// ---- POUs/IEC61850Server/WTURBINE/LD0/WTUR1/CDCs/FB_DO_WTURBINE_LD0_WTUR1_Beh.TcPOU
{attribute 'no_assign'}
FUNCTION_BLOCK FB_DO_WTURBINE_LD0_WTUR1_Beh EXTENDS FB_AcsiCommonDataClass
VAR_INPUT
	stVal: FB_AcsiDATypeBeh := (Fc:=ACSI_FC_ST, TrgOp:=ACSI_TrgOp_dchg OR ACSI_TrgOp_dupd, bLinkResult:=THIS^.AddDataToContainer(ipData:=stVal));
	q: FB_AcsiDATypeQuality := (Fc:=ACSI_FC_ST, TrgOp:=ACSI_TrgOp_qchg, bLinkResult:=THIS^.AddDataToContainer(ipData:=q));
	t: FB_AcsiDATypeTimeStamp := (Fc:=ACSI_FC_ST, bLinkResult:=THIS^.AddDataToContainer(ipData:=t));
END_VAR
VAR
END_VAR

END_FUNCTION_BLOCK

// ---- POUs/IEC61850Server/WTURBINE/LD0/WTUR1/CDCs/FB_DO_WTURBINE_LD0_WTUR1_TotWh.TcPOU
{attribute 'no_assign'}
FUNCTION_BLOCK FB_DO_WTURBINE_LD0_WTUR1_TotWh EXTENDS FB_AcsiCommonDataClass
VAR_INPUT
	cntVal: FB_DO_WTURBINE_LD0_WTUR1_TotWh_cntVal := (sClass:='BCR', bLinkResult:=THIS^.AddDataToContainer(ipData:=cntVal));
END_VAR
VAR
END_VAR

END_FUNCTION_BLOCK

// ---- POUs/IEC61850Server/WTURBINE/LD0/WTUR1/CDCs/FB_DO_WTURBINE_LD0_WTUR1_TotWh_cntVal.TcPOU
{attribute 'no_assign'}
FUNCTION_BLOCK FB_DO_WTURBINE_LD0_WTUR1_TotWh_cntVal EXTENDS FB_AcsiCommonDataClass
VAR_INPUT
	actVal: FB_AcsiBATypeINT64 := (Fc:=ACSI_FC_ST, TrgOp:=ACSI_TrgOp_dchg, bLinkResult:=THIS^.AddDataToContainer(ipData:=actVal));
	q: FB_AcsiDATypeQuality := (Fc:=ACSI_FC_ST, TrgOp:=ACSI_TrgOp_qchg, bLinkResult:=THIS^.AddDataToContainer(ipData:=q));
	t: FB_AcsiDATypeTimeStamp := (Fc:=ACSI_FC_ST, bLinkResult:=THIS^.AddDataToContainer(ipData:=t));
	pulsQty: FB_AcsiBATypeFLOAT32 := (Fc:=ACSI_FC_CF, TrgOp:=ACSI_TrgOp_dchg, bLinkResult:=THIS^.AddDataToContainer(ipData:=pulsQty));
END_VAR
VAR
END_VAR

END_FUNCTION_BLOCK

// ---- POUs/IEC61850Server/WTURBINE/LD0/WTUR1/CDCs/FB_DO_WTURBINE_LD0_WTUR1_TurSt.TcPOU
{attribute 'no_assign'}
FUNCTION_BLOCK FB_DO_WTURBINE_LD0_WTUR1_TurSt EXTENDS FB_AcsiCommonDataClass
VAR_INPUT
	st_: FB_DO_WTURBINE_LD0_WTUR1_TurSt_st := (sObjectName:='st', sClass:='ENS', bLinkResult:=THIS^.AddDataToContainer(ipData:=st_));
END_VAR
VAR
END_VAR

END_FUNCTION_BLOCK

// ---- POUs/IEC61850Server/WTURBINE/LD0/WTUR1/CDCs/FB_DO_WTURBINE_LD0_WTUR1_TurSt_st.TcPOU
{attribute 'no_assign'}
FUNCTION_BLOCK FB_DO_WTURBINE_LD0_WTUR1_TurSt_st EXTENDS FB_AcsiCommonDataClass
VAR_INPUT
	stVal: FB_AcsiDATypeTurSt := (Fc:=ACSI_FC_ST, TrgOp:=ACSI_TrgOp_dchg OR ACSI_TrgOp_dupd, bLinkResult:=THIS^.AddDataToContainer(ipData:=stVal));
	q: FB_AcsiDATypeQuality := (Fc:=ACSI_FC_ST, TrgOp:=ACSI_TrgOp_qchg, bLinkResult:=THIS^.AddDataToContainer(ipData:=q));
	t: FB_AcsiDATypeTimeStamp := (Fc:=ACSI_FC_ST, bLinkResult:=THIS^.AddDataToContainer(ipData:=t));
END_VAR
VAR
END_VAR

END_FUNCTION_BLOCK

// ---- POUs/IEC61850Server/WTURBINE/LD0/WTUR1/CDCs/FB_DO_WTURBINE_LD0_WTUR1_W.TcPOU
{attribute 'no_assign'}
FUNCTION_BLOCK FB_DO_WTURBINE_LD0_WTUR1_W EXTENDS FB_AcsiCommonDataClass
VAR_INPUT
	mag: FB_AcsiDATypeAnalogueValue := (Fc:=ACSI_FC_MX, TrgOp:=ACSI_TrgOp_dchg OR ACSI_TrgOp_dupd, i:=(bPresence:=FALSE), bLinkResult:=THIS^.AddDataToContainer(ipData:=mag));
	q: FB_AcsiDATypeQuality := (Fc:=ACSI_FC_MX, TrgOp:=ACSI_TrgOp_qchg, bLinkResult:=THIS^.AddDataToContainer(ipData:=q));
	t: FB_AcsiDATypeTimeStamp := (Fc:=ACSI_FC_MX, bLinkResult:=THIS^.AddDataToContainer(ipData:=t));
END_VAR
VAR
END_VAR

END_FUNCTION_BLOCK

// ---- POUs/IEC61850Server/WTURBINE/LD0/WTUR1/CDCs/FB_DO_WTURBINE_LD0_WTUR1_TurOp.TcPOU
{attribute 'no_assign'}
FUNCTION_BLOCK FB_DO_WTURBINE_LD0_WTUR1_TurOp EXTENDS FB_AcsiCommonDataClass
VAR_INPUT
	cmdAcs: FB_AcsiBATypeINT8U := (Fc:=ACSI_FC_CF, bLinkResult:=THIS^.AddDataToContainer(ipData:=cmdAcs));
	st_: FB_DO_WTURBINE_LD0_WTUR1_TurOp_st := (sObjectName:='st', sClass:='ENC', bLinkResult:=THIS^.AddDataToContainer(ipData:=st_));
END_VAR
VAR
END_VAR

END_FUNCTION_BLOCK

// ---- POUs/IEC61850Server/WTURBINE/LD0/WTUR1/CDCs/FB_DO_WTURBINE_LD0_WTUR1_TurOp_st.TcPOU
{attribute 'no_assign'}
FUNCTION_BLOCK FB_DO_WTURBINE_LD0_WTUR1_TurOp_st EXTENDS FB_AcsiCommonControllableDataClass
VAR_INPUT
	stVal: FB_AcsiDATypeTurOp := (Fc:=ACSI_FC_ST, TrgOp:=ACSI_TrgOp_dchg, bLinkResult:=THIS^.AddDataToContainer(ipData:=stVal));
	q: FB_AcsiDATypeQuality := (Fc:=ACSI_FC_ST, TrgOp:=ACSI_TrgOp_qchg, bLinkResult:=THIS^.AddDataToContainer(ipData:=q));
	t: FB_AcsiDATypeTimeStamp := (Fc:=ACSI_FC_ST, bLinkResult:=THIS^.AddDataToContainer(ipData:=t));
	ctlModel: FB_AcsiDATypeCtlModels := (Fc:=ACSI_FC_CF, TrgOp:=ACSI_TrgOp_dchg, eValue:=E_AcsiCtlModels.DirectWithNormalSecurity, bLinkResult:=THIS^.AddDataToContainer(ipData:=ctlModel));
	Cancel: FB_AcsiCDC_Cancel_ENUMERATED := (Fc:=ACSI_FC_CO, bLinkResult:=THIS^.AddDataToContainer(ipData:=Cancel));
	Oper: FB_AcsiCDC_Oper_ENUMERATED := (Fc:=ACSI_FC_CO, bLinkResult:=THIS^.AddDataToContainer(ipData:=Oper));
	SBO: FB_AcsiCDC_SBO := (Fc:=ACSI_FC_CO, bLinkResult:=THIS^.AddDataToContainer(ipData:=SBO));
	
	fbControl: FB_DirectControl := (ipCtrl:=THIS^.AddServerJob(ipEvent:=fbControl, ipCompletion:=fbControl));
END_VAR
VAR
END_VAR

END_FUNCTION_BLOCK

// ---- POUs/IEC61850Server/WTURBINE/LD0/WTUR1/CDCs/FB_DO_WTURBINE_LD0_WTUR1_DmdWSpt.TcPOU
{attribute 'no_assign'}
FUNCTION_BLOCK FB_DO_WTURBINE_LD0_WTUR1_DmdWSpt EXTENDS FB_AcsiCommonDataClass
VAR_INPUT
	val: FB_DO_WTURBINE_LD0_WTUR1_DmdWSpt_val := (sClass:='APC', bLinkResult:=THIS^.AddDataToContainer(ipData:=val));
END_VAR
VAR
END_VAR

END_FUNCTION_BLOCK

// ---- POUs/IEC61850Server/WTURBINE/LD0/WTUR1/CDCs/FB_DO_WTURBINE_LD0_WTUR1_DmdWSpt_val.TcPOU
{attribute 'no_assign'}
FUNCTION_BLOCK FB_DO_WTURBINE_LD0_WTUR1_DmdWSpt_val EXTENDS FB_AcsiCommonControllableDataClass
VAR_INPUT
	origin: FB_AcsiDATypeOriginator := (Fc:=ACSI_FC_MX, bLinkResult:=THIS^.AddDataToContainer(ipData:=origin));
	mxVal: FB_AcsiDATypeAnalogueValue := (Fc:=ACSI_FC_MX, TrgOp:=ACSI_TrgOp_dchg, i:=(bPresence:=FALSE), bLinkResult:=THIS^.AddDataToContainer(ipData:=mxVal));
	q: FB_AcsiDATypeQuality := (Fc:=ACSI_FC_MX, TrgOp:=ACSI_TrgOp_qchg, bLinkResult:=THIS^.AddDataToContainer(ipData:=q));
	t: FB_AcsiDATypeTimeStamp := (Fc:=ACSI_FC_MX, bLinkResult:=THIS^.AddDataToContainer(ipData:=t));
	ctlModel: FB_AcsiDATypeCtlModels := (Fc:=ACSI_FC_CF, TrgOp:=ACSI_TrgOp_dchg, eValue:=E_AcsiCtlModels.DirectWithNormalSecurity, bLinkResult:=THIS^.AddDataToContainer(ipData:=ctlModel));
	Oper: FB_AcsiCDC_Oper_AnalogueValue := (Fc:=ACSI_FC_CO, ctlVal:=(i:=(bPresence:=FALSE)), bLinkResult:=THIS^.AddDataToContainer(ipData:=Oper));
	SBO: FB_AcsiCDC_SBO := (Fc:=ACSI_FC_CO, bLinkResult:=THIS^.AddDataToContainer(ipData:=SBO));
	Cancel: FB_AcsiCDC_Cancel_AnalogueValue := (Fc:=ACSI_FC_CO, ctlVal:=(i:=(bPresence:=FALSE)), bLinkResult:=THIS^.AddDataToContainer(ipData:=Cancel));
	
	fbControl: FB_DirectControl := (ipCtrl:=THIS^.AddServerJob(ipEvent:=fbControl, ipCompletion:=fbControl));
// 	fbControl: FB_SboControl := (ipCtrl:=THIS^.AddServerJob(ipEvent:=fbControl, ipCompletion:=fbControl));
END_VAR
VAR
END_VAR

END_FUNCTION_BLOCK

// ---- POUs/IEC61850Server/WTURBINE/LD0/WTUR1/CDCs/FB_DO_WTURBINE_LD0_WTUR1_TurCtl.TcPOU
{attribute 'no_assign'}
FUNCTION_BLOCK FB_DO_WTURBINE_LD0_WTUR1_TurCtl EXTENDS FB_AcsiCommonDataClass
VAR_INPUT
	st_: FB_DO_WTURBINE_LD0_WTUR1_TurCtl_st := (sObjectName:='st', sClass:='ENC', bLinkResult:=THIS^.AddDataToContainer(ipData:=st_));
END_VAR
VAR
END_VAR

END_FUNCTION_BLOCK

// ---- POUs/IEC61850Server/WTURBINE/LD0/WTUR1/CDCs/FB_DO_WTURBINE_LD0_WTUR1_TurCtl_st.TcPOU
{attribute 'no_assign'}
FUNCTION_BLOCK FB_DO_WTURBINE_LD0_WTUR1_TurCtl_st EXTENDS FB_AcsiCommonControllableDataClass
VAR_INPUT
	//stVal: FB_AcsiBATypeEnumerated := (Fc:=ACSI_FC_ST, TrgOp:=ACSI_TrgOp_dchg, bLinkResult:=THIS^.AddDataToContainer(ipData:=stVal));
	stVal: FB_AcsiDATypeTurOp := (Fc:=ACSI_FC_ST, TrgOp:=ACSI_TrgOp_dchg, bLinkResult:=THIS^.AddDataToContainer(ipData:=stVal));
	q: FB_AcsiDATypeQuality := (Fc:=ACSI_FC_ST, TrgOp:=ACSI_TrgOp_qchg, bLinkResult:=THIS^.AddDataToContainer(ipData:=q));
	t: FB_AcsiDATypeTimeStamp := (Fc:=ACSI_FC_ST, bLinkResult:=THIS^.AddDataToContainer(ipData:=t));
	ctlModel: FB_AcsiDATypeCtlModels := (Fc:=ACSI_FC_CF, TrgOp:=ACSI_TrgOp_dchg, eValue:=E_AcsiCtlModels.DirectWithNormalSecurity, bLinkResult:=THIS^.AddDataToContainer(ipData:=ctlModel));
	Cancel: FB_AcsiCDC_Cancel_ENUMERATED := (Fc:=ACSI_FC_CO, bLinkResult:=THIS^.AddDataToContainer(ipData:=Cancel));
	Oper: FB_AcsiCDC_Oper_ENUMERATED := (Fc:=ACSI_FC_CO, bLinkResult:=THIS^.AddDataToContainer(ipData:=Oper));
	SBO: FB_AcsiCDC_SBO := (Fc:=ACSI_FC_CO, bLinkResult:=THIS^.AddDataToContainer(ipData:=SBO));
	
	fbControl: FB_DirectControl := (ipCtrl:=THIS^.AddServerJob(ipEvent:=fbControl, ipCompletion:=fbControl));
END_VAR
VAR
END_VAR

END_FUNCTION_BLOCK

// ---- POUs/IEC61850Server/WTURBINE/LD0/WROT1/FB_LN_WTURBINE_LD0_WROT1.TcPOU
{attribute 'no_assign'}
FUNCTION_BLOCK FB_LN_WTURBINE_LD0_WROT1 EXTENDS FB_AcsiCommonLogicalNodeClass
VAR_INPUT
	Beh: FB_DO_WTURBINE_LD0_WROT1_Beh := (sClass:='ENS', bLinkResult:=THIS^.AddDataToContainer(ipData:=Beh));
	RotSpd: FB_DO_WTURBINE_LD0_WROT1_RotSpd := (sClass:='MV', bLinkResult:=THIS^.AddDataToContainer(ipData:=RotSpd));
	BlPthAngTgt: FB_DO_WTURBINE_LD0_WROT1_BlPthAngTgt := (sClass:='MV', bLinkResult:=THIS^.AddDataToContainer(ipData:=BlPthAngTgt));
	BlPthAngVal: FB_DO_WTURBINE_LD0_WROT1_BlPthAngVal := (sClass:='MV', bLinkResult:=THIS^.AddDataToContainer(ipData:=BlPthAngVal));
END_VAR
VAR
END_VAR

END_FUNCTION_BLOCK

// ---- POUs/IEC61850Server/WTURBINE/LD0/WROT1/CDCs/FB_DO_WTURBINE_LD0_WROT1_Beh.TcPOU
{attribute 'no_assign'}
FUNCTION_BLOCK FB_DO_WTURBINE_LD0_WROT1_Beh EXTENDS FB_AcsiCommonDataClass
VAR_INPUT
	stVal: FB_AcsiDATypeBeh := (Fc:=ACSI_FC_ST, TrgOp:=ACSI_TrgOp_dchg OR ACSI_TrgOp_dupd, bLinkResult:=THIS^.AddDataToContainer(ipData:=stVal));
	q: FB_AcsiDATypeQuality := (Fc:=ACSI_FC_ST, TrgOp:=ACSI_TrgOp_qchg, bLinkResult:=THIS^.AddDataToContainer(ipData:=q));
	t: FB_AcsiDATypeTimeStamp := (Fc:=ACSI_FC_ST, bLinkResult:=THIS^.AddDataToContainer(ipData:=t));
END_VAR
VAR
END_VAR

END_FUNCTION_BLOCK

// ---- POUs/IEC61850Server/WTURBINE/LD0/WROT1/CDCs/FB_DO_WTURBINE_LD0_WROT1_RotSpd.TcPOU
{attribute 'no_assign'}
FUNCTION_BLOCK FB_DO_WTURBINE_LD0_WROT1_RotSpd EXTENDS FB_AcsiCommonDataClass
VAR_INPUT
	mag: FB_AcsiDATypeAnalogueValue := (Fc:=ACSI_FC_MX, TrgOp:=ACSI_TrgOp_dchg OR ACSI_TrgOp_dupd, i:=(bPresence:=FALSE), bLinkResult:=THIS^.AddDataToContainer(ipData:=mag));
	q: FB_AcsiDATypeQuality := (Fc:=ACSI_FC_MX, TrgOp:=ACSI_TrgOp_qchg, bLinkResult:=THIS^.AddDataToContainer(ipData:=q));
	t: FB_AcsiDATypeTimeStamp := (Fc:=ACSI_FC_MX, bLinkResult:=THIS^.AddDataToContainer(ipData:=t));
END_VAR
VAR
END_VAR

END_FUNCTION_BLOCK

// ---- POUs/IEC61850Server/WTURBINE/LD0/WROT1/CDCs/FB_DO_WTURBINE_LD0_WROT1_BlPthAngTgt.TcPOU
{attribute 'no_assign'}
FUNCTION_BLOCK FB_DO_WTURBINE_LD0_WROT1_BlPthAngTgt EXTENDS FB_AcsiCommonDataClass
VAR_INPUT
	mag: FB_AcsiDATypeAnalogueValue := (Fc:=ACSI_FC_MX, TrgOp:=ACSI_TrgOp_dchg OR ACSI_TrgOp_dupd, i:=(bPresence:=FALSE), bLinkResult:=THIS^.AddDataToContainer(ipData:=mag));
	q: FB_AcsiDATypeQuality := (Fc:=ACSI_FC_MX, TrgOp:=ACSI_TrgOp_qchg, bLinkResult:=THIS^.AddDataToContainer(ipData:=q));
	t: FB_AcsiDATypeTimeStamp := (Fc:=ACSI_FC_MX, bLinkResult:=THIS^.AddDataToContainer(ipData:=t));
END_VAR
VAR
END_VAR

END_FUNCTION_BLOCK

// ---- POUs/IEC61850Server/WTURBINE/LD0/WROT1/CDCs/FB_DO_WTURBINE_LD0_WROT1_BlPthAngVal.TcPOU
{attribute 'no_assign'}
FUNCTION_BLOCK FB_DO_WTURBINE_LD0_WROT1_BlPthAngVal EXTENDS FB_AcsiCommonDataClass
VAR_INPUT
	mag: FB_AcsiDATypeAnalogueValue := (Fc:=ACSI_FC_MX, TrgOp:=ACSI_TrgOp_dchg OR ACSI_TrgOp_dupd, i:=(bPresence:=FALSE), bLinkResult:=THIS^.AddDataToContainer(ipData:=mag));
	q: FB_AcsiDATypeQuality := (Fc:=ACSI_FC_MX, TrgOp:=ACSI_TrgOp_qchg, bLinkResult:=THIS^.AddDataToContainer(ipData:=q));
	t: FB_AcsiDATypeTimeStamp := (Fc:=ACSI_FC_MX, bLinkResult:=THIS^.AddDataToContainer(ipData:=t));
END_VAR
VAR
END_VAR

END_FUNCTION_BLOCK

// ---- POUs/IEC61850Server/WTURBINE/LD0/WCNV1/FB_LN_WTURBINE_LD0_WCNV1.TcPOU
{attribute 'no_assign'}
FUNCTION_BLOCK FB_LN_WTURBINE_LD0_WCNV1 EXTENDS FB_AcsiCommonLogicalNodeClass
VAR_INPUT
	Beh: FB_DO_WTURBINE_LD0_WCNV1_Beh := (sClass:='ENS', bLinkResult:=THIS^.AddDataToContainer(ipData:=Beh));
	Torq: FB_DO_WTURBINE_LD0_WCNV1_Torq := (sClass:='MV', bLinkResult:=THIS^.AddDataToContainer(ipData:=Torq));
END_VAR
VAR
END_VAR

END_FUNCTION_BLOCK

// ---- POUs/IEC61850Server/WTURBINE/LD0/WCNV1/CDCs/FB_DO_WTURBINE_LD0_WCNV1_Beh.TcPOU
{attribute 'no_assign'}
FUNCTION_BLOCK FB_DO_WTURBINE_LD0_WCNV1_Beh EXTENDS FB_AcsiCommonDataClass
VAR_INPUT
	stVal: FB_AcsiDATypeBeh := (Fc:=ACSI_FC_ST, TrgOp:=ACSI_TrgOp_dchg OR ACSI_TrgOp_dupd, bLinkResult:=THIS^.AddDataToContainer(ipData:=stVal));
	q: FB_AcsiDATypeQuality := (Fc:=ACSI_FC_ST, TrgOp:=ACSI_TrgOp_qchg, bLinkResult:=THIS^.AddDataToContainer(ipData:=q));
	t: FB_AcsiDATypeTimeStamp := (Fc:=ACSI_FC_ST, bLinkResult:=THIS^.AddDataToContainer(ipData:=t));
END_VAR
VAR
END_VAR

END_FUNCTION_BLOCK

// ---- POUs/IEC61850Server/WTURBINE/LD0/WCNV1/CDCs/FB_DO_WTURBINE_LD0_WCNV1_Torq.TcPOU
{attribute 'no_assign'}
FUNCTION_BLOCK FB_DO_WTURBINE_LD0_WCNV1_Torq EXTENDS FB_AcsiCommonDataClass
VAR_INPUT
	mag: FB_AcsiDATypeAnalogueValue := (Fc:=ACSI_FC_MX, TrgOp:=ACSI_TrgOp_dchg OR ACSI_TrgOp_dupd, i:=(bPresence:=FALSE), bLinkResult:=THIS^.AddDataToContainer(ipData:=mag));
	q: FB_AcsiDATypeQuality := (Fc:=ACSI_FC_MX, TrgOp:=ACSI_TrgOp_qchg, bLinkResult:=THIS^.AddDataToContainer(ipData:=q));
	t: FB_AcsiDATypeTimeStamp := (Fc:=ACSI_FC_MX, bLinkResult:=THIS^.AddDataToContainer(ipData:=t));
END_VAR
VAR
END_VAR

END_FUNCTION_BLOCK

// ---- POUs/IEC61850Server/WTURBINE/LD0/WMET1/FB_LN_WTURBINE_LD0_WMET1.TcPOU
{attribute 'no_assign'}
FUNCTION_BLOCK FB_LN_WTURBINE_LD0_WMET1 EXTENDS FB_AcsiCommonLogicalNodeClass
VAR_INPUT
	Beh: FB_DO_WTURBINE_LD0_WMET1_Beh := (sClass:='ENS', bLinkResult:=THIS^.AddDataToContainer(ipData:=Beh));
	HorWdDir: FB_DO_WTURBINE_LD0_WMET1_HorWdDir := (sClass:='MV', bLinkResult:=THIS^.AddDataToContainer(ipData:=HorWdDir));
	HorWdSpd: FB_DO_WTURBINE_LD0_WMET1_HorWdSpd := (sClass:='MV', bLinkResult:=THIS^.AddDataToContainer(ipData:=HorWdSpd));
END_VAR
VAR
END_VAR

END_FUNCTION_BLOCK

// ---- POUs/IEC61850Server/WTURBINE/LD0/WMET1/CDCs/FB_DO_WTURBINE_LD0_WMET1_Beh.TcPOU
{attribute 'no_assign'}
FUNCTION_BLOCK FB_DO_WTURBINE_LD0_WMET1_Beh EXTENDS FB_AcsiCommonDataClass
VAR_INPUT
	stVal: FB_AcsiDATypeBeh := (Fc:=ACSI_FC_ST, TrgOp:=ACSI_TrgOp_dchg OR ACSI_TrgOp_dupd, bLinkResult:=THIS^.AddDataToContainer(ipData:=stVal));
	q: FB_AcsiDATypeQuality := (Fc:=ACSI_FC_ST, TrgOp:=ACSI_TrgOp_qchg, bLinkResult:=THIS^.AddDataToContainer(ipData:=q));
	t: FB_AcsiDATypeTimeStamp := (Fc:=ACSI_FC_ST, bLinkResult:=THIS^.AddDataToContainer(ipData:=t));
END_VAR
VAR
END_VAR

END_FUNCTION_BLOCK

// ---- POUs/IEC61850Server/WTURBINE/LD0/WMET1/CDCs/FB_DO_WTURBINE_LD0_WMET1_HorWdDir.TcPOU
{attribute 'no_assign'}
FUNCTION_BLOCK FB_DO_WTURBINE_LD0_WMET1_HorWdDir EXTENDS FB_AcsiCommonDataClass
VAR_INPUT
	mag: FB_AcsiDATypeAnalogueValue := (Fc:=ACSI_FC_MX, TrgOp:=ACSI_TrgOp_dchg OR ACSI_TrgOp_dupd, i:=(bPresence:=FALSE), bLinkResult:=THIS^.AddDataToContainer(ipData:=mag));
	q: FB_AcsiDATypeQuality := (Fc:=ACSI_FC_MX, TrgOp:=ACSI_TrgOp_qchg, bLinkResult:=THIS^.AddDataToContainer(ipData:=q));
	t: FB_AcsiDATypeTimeStamp := (Fc:=ACSI_FC_MX, bLinkResult:=THIS^.AddDataToContainer(ipData:=t));
END_VAR
VAR
END_VAR

END_FUNCTION_BLOCK

// ---- POUs/IEC61850Server/WTURBINE/LD0/WMET1/CDCs/FB_DO_WTURBINE_LD0_WMET1_HorWdSpd.TcPOU
{attribute 'no_assign'}
FUNCTION_BLOCK FB_DO_WTURBINE_LD0_WMET1_HorWdSpd EXTENDS FB_AcsiCommonDataClass
VAR_INPUT
	mag: FB_AcsiDATypeAnalogueValue := (Fc:=ACSI_FC_MX, TrgOp:=ACSI_TrgOp_dchg OR ACSI_TrgOp_dupd, i:=(bPresence:=FALSE), bLinkResult:=THIS^.AddDataToContainer(ipData:=mag));
	q: FB_AcsiDATypeQuality := (Fc:=ACSI_FC_MX, TrgOp:=ACSI_TrgOp_qchg, bLinkResult:=THIS^.AddDataToContainer(ipData:=q));
	t: FB_AcsiDATypeTimeStamp := (Fc:=ACSI_FC_MX, bLinkResult:=THIS^.AddDataToContainer(ipData:=t));
END_VAR
VAR
END_VAR

END_FUNCTION_BLOCK

// ---- POUs/IEC61850Server/WTURBINE/LD0/WALM1/FB_LN_WTURBINE_LD0_WALM1.TcPOU
{attribute 'no_assign'}
FUNCTION_BLOCK FB_LN_WTURBINE_LD0_WALM1 EXTENDS FB_AcsiCommonLogicalNodeClass
VAR_INPUT
	Beh: FB_DO_WTURBINE_LD0_WALM1_Beh := (sClass:='ENS', bLinkResult:=THIS^.AddDataToContainer(ipData:=Beh));
END_VAR
VAR
END_VAR

END_FUNCTION_BLOCK

// ---- POUs/IEC61850Server/WTURBINE/LD0/WALM1/CDCs/FB_DO_WTURBINE_LD0_WALM1_Beh.TcPOU
{attribute 'no_assign'}
FUNCTION_BLOCK FB_DO_WTURBINE_LD0_WALM1_Beh EXTENDS FB_AcsiCommonDataClass
VAR_INPUT
	stVal: FB_AcsiDATypeBeh := (Fc:=ACSI_FC_ST, TrgOp:=ACSI_TrgOp_dchg OR ACSI_TrgOp_dupd, bLinkResult:=THIS^.AddDataToContainer(ipData:=stVal));
	q: FB_AcsiDATypeQuality := (Fc:=ACSI_FC_ST, TrgOp:=ACSI_TrgOp_qchg, bLinkResult:=THIS^.AddDataToContainer(ipData:=q));
	t: FB_AcsiDATypeTimeStamp := (Fc:=ACSI_FC_ST, bLinkResult:=THIS^.AddDataToContainer(ipData:=t));
END_VAR
VAR
END_VAR

END_FUNCTION_BLOCK

// ---- POUs/IEC61850Server/WTURBINE/LD0/WYAW1/FB_LN_WTURBINE_LD0_WYAW1.TcPOU
{attribute 'no_assign'}
FUNCTION_BLOCK FB_LN_WTURBINE_LD0_WYAW1 EXTENDS FB_AcsiCommonLogicalNodeClass
VAR_INPUT
	Beh: FB_DO_WTURBINE_LD0_WYAW1_Beh := (sClass:='ENS', bLinkResult:=THIS^.AddDataToContainer(ipData:=Beh));
	YwAng: FB_DO_WTURBINE_LD0_WYAW1_YwAng := (sClass:='MV', bLinkResult:=THIS^.AddDataToContainer(ipData:=YwAng));
	CabWup: FB_DO_WTURBINE_LD0_WYAW1_CabWup := (sClass:='MV', bLinkResult:=THIS^.AddDataToContainer(ipData:=CabWup));
	YwAngSpt: FB_DO_WTURBINE_LD0_WYAW1_YwAngSpt := (sClass:='SPV', bLinkResult:=THIS^.AddDataToContainer(ipData:=YwAngSpt));
END_VAR
VAR
END_VAR

END_FUNCTION_BLOCK

// ---- POUs/IEC61850Server/WTURBINE/LD0/WYAW1/CDCs/FB_DO_WTURBINE_LD0_WYAW1_Beh.TcPOU
{attribute 'no_assign'}
FUNCTION_BLOCK FB_DO_WTURBINE_LD0_WYAW1_Beh EXTENDS FB_AcsiCommonDataClass
VAR_INPUT
	stVal: FB_AcsiDATypeBeh := (Fc:=ACSI_FC_ST, TrgOp:=ACSI_TrgOp_dchg OR ACSI_TrgOp_dupd, bLinkResult:=THIS^.AddDataToContainer(ipData:=stVal));
	q: FB_AcsiDATypeQuality := (Fc:=ACSI_FC_ST, TrgOp:=ACSI_TrgOp_qchg, bLinkResult:=THIS^.AddDataToContainer(ipData:=q));
	t: FB_AcsiDATypeTimeStamp := (Fc:=ACSI_FC_ST, bLinkResult:=THIS^.AddDataToContainer(ipData:=t));
END_VAR
VAR
END_VAR

END_FUNCTION_BLOCK

// ---- POUs/IEC61850Server/WTURBINE/LD0/WYAW1/CDCs/FB_DO_WTURBINE_LD0_WYAW1_YwAng.TcPOU
{attribute 'no_assign'}
FUNCTION_BLOCK FB_DO_WTURBINE_LD0_WYAW1_YwAng EXTENDS FB_AcsiCommonDataClass
VAR_INPUT
	mag: FB_AcsiDATypeAnalogueValue := (Fc:=ACSI_FC_MX, TrgOp:=ACSI_TrgOp_dchg OR ACSI_TrgOp_dupd, i:=(bPresence:=FALSE), bLinkResult:=THIS^.AddDataToContainer(ipData:=mag));
	q: FB_AcsiDATypeQuality := (Fc:=ACSI_FC_MX, TrgOp:=ACSI_TrgOp_qchg, bLinkResult:=THIS^.AddDataToContainer(ipData:=q));
	t: FB_AcsiDATypeTimeStamp := (Fc:=ACSI_FC_MX, bLinkResult:=THIS^.AddDataToContainer(ipData:=t));
END_VAR
VAR
END_VAR

END_FUNCTION_BLOCK

// ---- POUs/IEC61850Server/WTURBINE/LD0/WYAW1/CDCs/FB_DO_WTURBINE_LD0_WYAW1_CabWup.TcPOU
{attribute 'no_assign'}
FUNCTION_BLOCK FB_DO_WTURBINE_LD0_WYAW1_CabWup EXTENDS FB_AcsiCommonDataClass
VAR_INPUT
	mag: FB_AcsiDATypeAnalogueValue := (Fc:=ACSI_FC_MX, TrgOp:=ACSI_TrgOp_dchg OR ACSI_TrgOp_dupd, i:=(bPresence:=FALSE), f:=(bPresence:=FALSE), bLinkResult:=THIS^.AddDataToContainer(ipData:=mag));
	q: FB_AcsiDATypeQuality := (Fc:=ACSI_FC_MX, TrgOp:=ACSI_TrgOp_qchg, bLinkResult:=THIS^.AddDataToContainer(ipData:=q));
	t: FB_AcsiDATypeTimeStamp := (Fc:=ACSI_FC_MX, bLinkResult:=THIS^.AddDataToContainer(ipData:=t));
END_VAR
VAR
END_VAR

END_FUNCTION_BLOCK

// ---- POUs/IEC61850Server/WTURBINE/LD0/WYAW1/CDCs/FB_DO_WTURBINE_LD0_WYAW1_YwAngSpt.TcPOU
{attribute 'no_assign'}
FUNCTION_BLOCK FB_DO_WTURBINE_LD0_WYAW1_YwAngSpt EXTENDS FB_AcsiCommonDataClass
VAR_INPUT
	val: FB_DO_WTURBINE_LD0_WYAW1_YwAngSpt_val := (sClass:='APC', bLinkResult:=THIS^.AddDataToContainer(ipData:=val));
END_VAR
VAR
END_VAR

END_FUNCTION_BLOCK

// ---- POUs/IEC61850Server/WTURBINE/LD0/WYAW1/CDCs/FB_DO_WTURBINE_LD0_WYAW1_YwAngSpt_val.TcPOU
{attribute 'no_assign'}
FUNCTION_BLOCK FB_DO_WTURBINE_LD0_WYAW1_YwAngSpt_val EXTENDS FB_AcsiCommonControllableDataClass
VAR_INPUT
	origin: FB_AcsiDATypeOriginator := (Fc:=ACSI_FC_MX, bLinkResult:=THIS^.AddDataToContainer(ipData:=origin));
	mxVal: FB_AcsiDATypeAnalogueValue := (Fc:=ACSI_FC_MX, TrgOp:=ACSI_TrgOp_dchg, i:=(bPresence:=FALSE), bLinkResult:=THIS^.AddDataToContainer(ipData:=mxVal));
	q: FB_AcsiDATypeQuality := (Fc:=ACSI_FC_MX, TrgOp:=ACSI_TrgOp_qchg, bLinkResult:=THIS^.AddDataToContainer(ipData:=q));
	t: FB_AcsiDATypeTimeStamp := (Fc:=ACSI_FC_MX, bLinkResult:=THIS^.AddDataToContainer(ipData:=t));
	ctlModel: FB_AcsiDATypeCtlModels := (Fc:=ACSI_FC_CF, TrgOp:=ACSI_TrgOp_dchg, eValue:=E_AcsiCtlModels.DirectWithNormalSecurity, bLinkResult:=THIS^.AddDataToContainer(ipData:=ctlModel));
	Oper: FB_AcsiCDC_Oper_AnalogueValue := (Fc:=ACSI_FC_CO, ctlVal:=(i:=(bPresence:=FALSE)), bLinkResult:=THIS^.AddDataToContainer(ipData:=Oper));
	
	fbControl: FB_DirectControl := (ipCtrl:=THIS^.AddServerJob(ipEvent:=fbControl, ipCompletion:=fbControl));
END_VAR
VAR
END_VAR

END_FUNCTION_BLOCK

// ---- POUs/IEC61850Server/WTURBINE/LD0/WPPD1/FB_LN_WTURBINE_LD0_WPPD1.TcPOU
{attribute 'no_assign'}
FUNCTION_BLOCK FB_LN_WTURBINE_LD0_WPPD1 EXTENDS FB_AcsiCommonLogicalNodeClass
VAR_INPUT
	Beh: FB_DO_WTURBINE_LD0_WPPD1_Beh := (sClass:='ENS', bLinkResult:=THIS^.AddDataToContainer(ipData:=Beh));
	DevSt: FB_DO_WTURBINE_LD0_WPPD1_DevSt := (sClass:='STV', bLinkResult:=THIS^.AddDataToContainer(ipData:=DevSt));
	DevOp: FB_DO_WTURBINE_LD0_WPPD1_DevOp := (sClass:='CMD', bLinkResult:=THIS^.AddDataToContainer(ipData:=DevOp));
	ClrOp: FB_DO_WTURBINE_LD0_WPPD1_ClrOp := (sClass:='CMD', bLinkResult:=THIS^.AddDataToContainer(ipData:=ClrOp));
	
	ds01: FB_DS_TEMPLATE_LD1_WPPD1_ds01 := (bLinkResult:=THIS^.AddDataSetToContainer(ipDataSet:=ds01));
	
	urcb01: FB_ScsmUrCBImplClass := (RptID:=(sValue:='WTURBINELD0/WPPD1.urcb01'), DatSet:=(sValue:='WTURBINELD0/WPPD1.ds01'), OptFlds:=(SequenceNumber:=FALSE, ReportTimeStamp:=FALSE, ReasonForInclusion:=FALSE, DataSetName:=FALSE, DataReference:=FALSE, BufferOverflow:=FALSE, EntryID:=FALSE, ConfRevision:=FALSE), TrgOps:=(DataChange:=FALSE, QualityChange:=FALSE, DataUpdate:=FALSE, Integrity:=FALSE, GeneralInterrogation:=TRUE), bLinkResult:=THIS^.AddUnbufferedReportControlBlockToContainer(ipUnbufferedReportControlBlock:=urcb01));
END_VAR
VAR
END_VAR

END_FUNCTION_BLOCK

// ---- POUs/IEC61850Server/WTURBINE/LD0/WPPD1/CDCs/FB_DO_WTURBINE_LD0_WPPD1_Beh.TcPOU
{attribute 'no_assign'}
FUNCTION_BLOCK FB_DO_WTURBINE_LD0_WPPD1_Beh EXTENDS FB_AcsiCommonDataClass
VAR_INPUT
	stVal: FB_AcsiDATypeBeh := (Fc:=ACSI_FC_ST, TrgOp:=ACSI_TrgOp_dchg OR ACSI_TrgOp_dupd, bLinkResult:=THIS^.AddDataToContainer(ipData:=stVal));
	q: FB_AcsiDATypeQuality := (Fc:=ACSI_FC_ST, TrgOp:=ACSI_TrgOp_qchg, bLinkResult:=THIS^.AddDataToContainer(ipData:=q));
	t: FB_AcsiDATypeTimeStamp := (Fc:=ACSI_FC_ST, bLinkResult:=THIS^.AddDataToContainer(ipData:=t));
END_VAR
VAR
END_VAR

END_FUNCTION_BLOCK

// ---- POUs/IEC61850Server/WTURBINE/LD0/WPPD1/CDCs/FB_DO_WTURBINE_LD0_WPPD1_DevSt.TcPOU
{attribute 'no_assign'}
FUNCTION_BLOCK FB_DO_WTURBINE_LD0_WPPD1_DevSt EXTENDS FB_AcsiCommonDataClass
VAR_INPUT
	st_: FB_DO_WTURBINE_LD0_WPPD1_DevSt_st := (sObjectName:='st', sClass:='ENS', bLinkResult:=THIS^.AddDataToContainer(ipData:=st_));
END_VAR
VAR
END_VAR

END_FUNCTION_BLOCK

// ---- POUs/IEC61850Server/WTURBINE/LD0/WPPD1/CDCs/FB_DO_WTURBINE_LD0_WPPD1_DevSt_st.TcPOU
{attribute 'no_assign'}
FUNCTION_BLOCK FB_DO_WTURBINE_LD0_WPPD1_DevSt_st EXTENDS FB_AcsiCommonDataClass
VAR_INPUT
	stVal: FB_AcsiDATypeDevSt := (Fc:=ACSI_FC_ST, TrgOp:=ACSI_TrgOp_dchg OR ACSI_TrgOp_dupd, bLinkResult:=THIS^.AddDataToContainer(ipData:=stVal));
	q: FB_AcsiDATypeQuality := (Fc:=ACSI_FC_ST, TrgOp:=ACSI_TrgOp_qchg, bLinkResult:=THIS^.AddDataToContainer(ipData:=q));
	t: FB_AcsiDATypeTimeStamp := (Fc:=ACSI_FC_ST, bLinkResult:=THIS^.AddDataToContainer(ipData:=t));
END_VAR
VAR
END_VAR

END_FUNCTION_BLOCK

// ---- POUs/IEC61850Server/WTURBINE/LD0/WPPD1/CDCs/FB_DO_WTURBINE_LD0_WPPD1_DevOp.TcPOU
{attribute 'no_assign'}
FUNCTION_BLOCK FB_DO_WTURBINE_LD0_WPPD1_DevOp EXTENDS FB_AcsiCommonDataClass
VAR_INPUT
	st_: FB_DO_WTURBINE_LD0_WPPD1_DevOp_st := (sObjectName:='st', sClass:='ENC', bLinkResult:=THIS^.AddDataToContainer(ipData:=st_));
END_VAR
VAR
END_VAR

END_FUNCTION_BLOCK

// ---- POUs/IEC61850Server/WTURBINE/LD0/WPPD1/CDCs/FB_DO_WTURBINE_LD0_WPPD1_DevOp_st.TcPOU
{attribute 'no_assign'}
FUNCTION_BLOCK FB_DO_WTURBINE_LD0_WPPD1_DevOp_st EXTENDS FB_AcsiCommonControllableDataClass
VAR_INPUT
	origin: FB_AcsiDATypeOriginator := (Fc:=ACSI_FC_ST, bLinkResult:=THIS^.AddDataToContainer(ipData:=origin));
	stVal: FB_AcsiDATypeDevOp := (Fc:=ACSI_FC_ST, TrgOp:=ACSI_TrgOp_dchg, bLinkResult:=THIS^.AddDataToContainer(ipData:=stVal));
	q: FB_AcsiDATypeQuality := (Fc:=ACSI_FC_ST, TrgOp:=ACSI_TrgOp_qchg, bLinkResult:=THIS^.AddDataToContainer(ipData:=q));
	t: FB_AcsiDATypeTimeStamp := (Fc:=ACSI_FC_ST, bLinkResult:=THIS^.AddDataToContainer(ipData:=t));
	ctlModel: FB_AcsiDATypeCtlModels := (Fc:=ACSI_FC_CF, TrgOp:=ACSI_TrgOp_dchg, bLinkResult:=THIS^.AddDataToContainer(ipData:=ctlModel));
	Cancel: FB_AcsiDATypeDelAct := (Fc:=ACSI_FC_CO, bLinkResult:=THIS^.AddDataToContainer(ipData:=Cancel));
	Oper: FB_AcsiCDC_Oper_ENUMERATED := (Fc:=ACSI_FC_CO, bLinkResult:=THIS^.AddDataToContainer(ipData:=Oper));
	SBO: FB_AcsiCDC_SBO := (Fc:=ACSI_FC_CO, bLinkResult:=THIS^.AddDataToContainer(ipData:=SBO));
	
	fbControl: FB_DirectControl := (ipCtrl:=THIS^.AddServerJob(ipEvent:=fbControl, ipCompletion:=fbControl));
END_VAR
VAR
END_VAR

END_FUNCTION_BLOCK

// ---- POUs/IEC61850Server/WTURBINE/LD0/WPPD1/CDCs/FB_DO_WTURBINE_LD0_WPPD1_ClrOp.TcPOU
{attribute 'no_assign'}
FUNCTION_BLOCK FB_DO_WTURBINE_LD0_WPPD1_ClrOp EXTENDS FB_AcsiCommonDataClass
VAR_INPUT
	st_: FB_DO_WTURBINE_LD0_WPPD1_ClrOp_st := (sObjectName:='st', sClass:='ENC', bLinkResult:=THIS^.AddDataToContainer(ipData:=st_));
END_VAR
VAR
END_VAR

END_FUNCTION_BLOCK

// ---- POUs/IEC61850Server/WTURBINE/LD0/WPPD1/CDCs/FB_DO_WTURBINE_LD0_WPPD1_ClrOp_st.TcPOU
{attribute 'no_assign'}
FUNCTION_BLOCK FB_DO_WTURBINE_LD0_WPPD1_ClrOp_st EXTENDS FB_AcsiCommonControllableDataClass
VAR_INPUT
	stVal: FB_AcsiBATypeENUMERATED := (Fc:=ACSI_FC_ST, TrgOp:=ACSI_TrgOp_dchg, bLinkResult:=THIS^.AddDataToContainer(ipData:=stVal));
	q: FB_AcsiDATypeQuality := (Fc:=ACSI_FC_ST, TrgOp:=ACSI_TrgOp_qchg, bLinkResult:=THIS^.AddDataToContainer(ipData:=q));
	t: FB_AcsiDATypeTimeStamp := (Fc:=ACSI_FC_ST, bLinkResult:=THIS^.AddDataToContainer(ipData:=t));
	ctlModel: FB_AcsiDATypeCtlModels := (Fc:=ACSI_FC_CF, TrgOp:=ACSI_TrgOp_dchg, bLinkResult:=THIS^.AddDataToContainer(ipData:=ctlModel));
	Cancel: FB_AcsiCDC_Cancel_ENUMERATED := (Fc:=ACSI_FC_CO, bLinkResult:=THIS^.AddDataToContainer(ipData:=Cancel));
	Oper: FB_AcsiCDC_Oper_ENUMERATED := (Fc:=ACSI_FC_CO, bLinkResult:=THIS^.AddDataToContainer(ipData:=Oper));
	SBO: FB_AcsiCDC_SBO := (Fc:=ACSI_FC_CO, bLinkResult:=THIS^.AddDataToContainer(ipData:=SBO));
	
	fbControl: FB_DirectControl := (ipCtrl:=THIS^.AddServerJob(ipEvent:=fbControl, ipCompletion:=fbControl));
END_VAR
VAR
END_VAR

END_FUNCTION_BLOCK

// ---- POUs/IEC61850Server/WTURBINE/LD0/WPPD1/DataSets/FB_DS_TEMPLATE_LD1_WPPD1_ds01.TcPOU
{attribute 'no_assign'}
{attribute 'call_after_init'}
FUNCTION_BLOCK FB_DS_TEMPLATE_LD1_WPPD1_ds01 EXTENDS FB_AcsiCommonDataSetClass
VAR
END_VAR

METHOD OnInit : BOOL
VAR
	nID : UDINT;
	i : UDINT;
END_VAR
// First find the nID this is part of
nID := c_nNumTurbines + 10;
FOR i := 1 TO c_nNumTurbines DO
    IF ADR(fbWTURBINE[i].WTURBINELD0.WPPD1.ds01) = ADR(THIS^) THEN
        nID := i;
        EXIT;
    END_IF
END_FOR

IF NOT DeleteAllMembers() THEN RETURN; END_IF
IF NOT AddMember(ipData:=fbWTURBINE[nID].WTURBINELD0.WYAW1.YwAng, eFc:=E_AcsiFc.MX) THEN RETURN; END_IF
IF NOT AddMember(ipData:=fbWTURBINE[nID].WTURBINELD0.WTUR1.W, eFc:=E_AcsiFc.MX) THEN RETURN; END_IF
IF NOT AddMember(ipData:=fbWTURBINE[nID].WTURBINELD0.WROT1.RotSpd, eFc:=E_AcsiFc.MX) THEN RETURN; END_IF
IF NOT AddMember(ipData:=fbWTURBINE[nID].WTURBINELD0.WROT1.BlPthAngTgt, eFc:=E_AcsiFc.MX) THEN RETURN; END_IF
IF NOT AddMember(ipData:=fbWTURBINE[nID].WTURBINELD0.WROT1.BlPthAngVal, eFc:=E_AcsiFc.MX) THEN RETURN; END_IF
IF NOT AddMember(ipData:=fbWTURBINE[nID].WTURBINELD0.WMET1.HorWdDir, eFc:=E_AcsiFc.MX) THEN RETURN; END_IF
IF NOT AddMember(ipData:=fbWTURBINE[nID].WTURBINELD0.WMET1.HorWdSpd, eFc:=E_AcsiFc.MX) THEN RETURN; END_IF
IF NOT AddMember(ipData:=fbWTURBINE[nID].WTURBINELD0.WCNV1.Torq, eFc:=E_AcsiFc.MX) THEN RETURN; END_IF
OnInit:= TRUE;
END_METHOD

END_FUNCTION_BLOCK

// ---- POUs/IEC61850Server/FB_WTURBINEServerSession.TcPOU
{attribute 'no_assign'}
FUNCTION_BLOCK FB_WTURBINEServerSession IMPLEMENTS I_ScsmAbortIndEventSink, I_ScsmAssociateIndEventSink, I_ScsmReleaseIndEventSink
VAR_INPUT
	fbConnection		: FB_iec61850ConnectionClass := (ipAbortInd:=THIS^, ipAssociateInd:=THIS^, ipReleaseInd:=THIS^);
	nID					: UDINT;
END_VAR
VAR
	_bAbort				: BOOL; (* Rising edge activates AbortReq() command execution *)
	_bDisconnect		: BOOL; (* Rising edge activates ReleaseReq() command execution *)
	
	state				: BYTE;
	eState				: E_AsyncEnvironmentState; (* Environment state *)
	eLinkStatus			: E_ScsmLinkStatus; (* Network adapter link status *)
	bBusy				: BOOL; (* If TRUE => command execution is busy *)
	bSuccess			: BOOL;
	ipResult			: I_AsyncServiceResultClass;
	sLastErrorResult	: T_MaxString;
	fbAbortReason		: FB_ServiceErrorClass := (stError:=SUCCESS_EVENT);
	sLastAbortReason	: T_MaxString;
END_VAR

fbConnection.Execute();
eState:= fbConnection.eState;
eLinkStatus:= fbConnection.eLinkStatus;

(* Execute control model control block implementations *)
// fbWTURBINE.WTURBINELD0.LLN0.Mod_.fbControl.Execute();
// fbWTURBINE.WTURBINELD0.WTUR1.CmdBlk.fbControl.Execute();
// fbWTURBINE.WTURBINELD0.WNAC1.CtlMd.fbControl.Execute();
// fbWTURBINE.WTURBINELD0.WYAW1.YwBrk.fbControl.Execute();

// fbWTURBINE[nID].WTURBINELD0.LLN0.Mod_.fbControl.Execute();
// fbWTURBINE[nID].WTURBINELD0.WTUR1.CmdBlk.fbControl.Execute();
// fbWTURBINE[nID].WTURBINELD0.WNAC1.CtlMd.fbControl.Execute();
// fbWTURBINE[nID].WTURBINELD0.WYAW1.YwBrk.fbControl.Execute();
// fbWTURBINE[nID].WTURBINELD0.WTUR1.DmdWSpt.fbControl.Execute();

(* Execute server control block implementations *)
fbWTURBINE[nID].WTURBINELD0.WPPD1.urcb01.Server.Execute();

fbWTURBINE[nID].WTURBINELD0.LLN0.Mod_.fbControl.Execute();
fbWTURBINE[nID].WTURBINELD0.WTUR1.TurOp.st_.fbControl.Execute();
fbWTURBINE[nID].WTURBINELD0.WTUR1.TurCtl.st_.fbControl.Execute();
fbWTURBINE[nID].WTURBINELD0.WTUR1.DmdWSpt.val.fbControl.Execute();
fbWTURBINE[nID].WTURBINELD0.WYAW1.YwAngSpt.val.fbControl.Execute();
fbWTURBINE[nID].WTURBINELD0.WPPD1.DevOp.st_.fbControl.Execute();
fbWTURBINE[nID].WTURBINELD0.WPPD1.ClrOp.st_.fbControl.Execute();

CASE state OF
	0: (* Initial state *)
		IF _bAbort THEN (* Abort connection => execute AbortReq() command *)
			_bAbort:= FALSE;
			bSuccess:= fbConnection.AbortReq(ipReason:=fbAbortReason, ipSink:=0, ipResult=>ipResult);
			state:= SEL(bSuccess, 100, 1);
		ELSIF eState = E_AsyncEnvironmentState.Established AND _bDisconnect THEN (* Close/release connection => execute ReleaseReq() command *)
			_bDisconnect:= FALSE;
			bSuccess:= fbConnection.ReleaseReq(ipSink:=0, ipResult=>ipResult);
			state:= SEL(bSuccess, 100, 1);
		ELSIF eState = E_AsyncEnvironmentState.Established THEN (* Connection established => exchange IED data *)
			state:= 10;
		END_IF
		_bDisconnect:= FALSE;
		(*==================================================================================================================================================================*)
	1: (* Wait for AbortReq() or ReleaseReq() command completion *)
		IF ipResult <> 0 THEN
			ipResult.Execute();
			IF NOT (bBusy:=ipResult.IsBusy()) THEN
				state:= SEL(ipResult.IsCompleted(), 100(* failed or aborted *), 0(* succeeded *));
			END_IF
		END_IF
		(*==================================================================================================================================================================*)
	10: (* connection established *)
		state:= 0;
		(*==================================================================================================================================================================*)
	100: (* Error state *)
		state:= 0;
		IF ipResult <> 0 THEN
			sLastErrorResult:= ipResult.Dump();
		END_IF
END_CASE

PROPERTY bAbort : BOOL
SET
_bAbort:= bAbort;
END_SET
END_PROPERTY

PROPERTY bDisconnect : BOOL
SET
_bDisconnect:= bDisconnect;
END_SET
END_PROPERTY

(* This method receives IEC61850::Abort.ind primitive. *)
METHOD OnAbortInd
VAR_INPUT
	ipAA		: I_ScsmAssociationClass; (* Application association. If = 0 => optional. *)
	bPAbort		: BOOL; (* TRUE => P-Abort.request(), issued by provider, FALSE => Abort.request(), issued by user. *)
	ipReason	: I_ServiceErrorClass; (* Abort reason. *)
	ipData		: I_BaseStreamClass; (* Optional data. If = 0 => default, no data. *)
END_VAR
VAR
END_VAR
IF ipReason <> 0 THEN
	sLastAbortReason:= ipReason.Dump();
END_IF
END_METHOD

(* This method receives IEC61850::Associate.ind primitive. *)
METHOD OnAssociateInd : BOOL
VAR_INPUT
	ipAA			: I_ScsmAssociationClass; (* Application association. If = 0 => optional. *)
END_VAR
VAR_OUTPUT
	ipResult		: I_AsyncServiceResultClass; (* Interface pointer to service state and result information *)
END_VAR
VAR
END_VAR
sLastAbortReason:= '';
sLastErrorResult:= '';
OnAssociateInd:= fbConnection.AssociateRsp(ipResult=>ipResult);
END_METHOD

(* This method receives IEC61850::Release.ind primitive. *)
METHOD OnReleaseInd : BOOL
VAR_INPUT
	ipAA	: I_ScsmAssociationClass; (* Application association. If = 0 => optional. *)
END_VAR
VAR_OUTPUT
	ipResult: I_AsyncServiceResultClass;
END_VAR
VAR
END_VAR
OnReleaseInd:= fbConnection.ReleaseRsp(ipResult=>ipResult);
END_METHOD

END_FUNCTION_BLOCK

// ---- POUs/IEC61850Server/FB_WTURBINEGse.TcPOU
{attribute 'no_assign'}
FUNCTION_BLOCK FB_WTURBINEGse IMPLEMENTS I_GseLinkStatusEventSink
VAR_INPUT
	fbAdapter		: FB_GseAdapterClass := (ipLinkStatus:=THIS^);
END_VAR
VAR
	eLinkStatus		: E_GseLinkStatus;
	
	bSuccess		: BOOL;
	ipError			: I_ServiceErrorClass;
	
	bStart			: BOOL := TRUE; (* Rising edge starts publishing of GOOSE data *)
	bStop			: BOOL; (* Rising edge stops publishing of GOOSE data *)
	bUpdate			: BOOL; (* Rising edge updates published GOOSE data *)
END_VAR

(*=========================================================================================*)
bSuccess:= fbAdapter.Execute(ipError=>ipError); (* Execute network adapter *)

(*=========================================================================================*)
// IF bStart THEN (* Start publishing of GOOSE data *)
// 	bStart:= FALSE;
// 	bSuccess:= fbWTURBINE.WTURBINELD0.LLN0.gocb01.Publisher.Start(ipAdapter:=fbAdapter, ipError=>ipError);
// ELSIF bStop THEN (* Stop publishing of GOOSE data *)
// 	bStop:= FALSE;
// 	bSuccess:= fbWTURBINE.WTURBINELD0.LLN0.gocb01.Publisher.Stop(ipError=>ipError);
// ELSIF bUpdate THEN (* Update published GOOSE data *)
// 	bUpdate:= FALSE;
// 	bSuccess:= fbWTURBINE.WTURBINELD0.LLN0.gocb01.Publisher.Update(ipError=>ipError);
// ELSE (* Execute publisher GoCB's *)
// 	bSuccess:= fbWTURBINE.WTURBINELD0.LLN0.gocb01.Publisher.Execute(ipError=>ipError);
// END_IF

(* This method is called every time the network adapter link status changes. *)
METHOD OnLinkStatusChange
VAR_INPUT
	ipAdapter	: I_GseAdapterClass;
	eStatus		: E_GseLinkStatus;
END_VAR
VAR
END_VAR
eLinkStatus:= eStatus;
END_METHOD

END_FUNCTION_BLOCK

// ---- POUs/IEC61850Server/FB_DirectControlEnhanced.TcPOU
FUNCTION_BLOCK FB_DirectControlEnhanced EXTENDS FB_DirectControl
VAR
END_VAR

METHOD Execute : BOOL
VAR
	bTestOk: BOOL; (*Used to cache the return value of the last '_OperativeTest' or '_DynamicTest' method call*)
	eError: E_AcsiServiceError; (*Used to cache the returned error of the last '_OperativeTest' or '_DynamicTest' method call*)
	tValue: T_UtcTime; (*Used to cache the current system time for 'tOpOk'*)
END_VAR
IF (_ipCtrl <> 0) AND_THEN (_ipCtrl.ipOper <> 0) THEN
	(* Initialize function block in the first cycle *)
	IF NOT bInit THEN
		_Init();
		bInit:=TRUE;
	END_IF

	CASE _eControlState OF
		E_DirectControlState.Ready:
			(* Check if ControlState changed in the last cycle *)
			IF bNewState THEN
				bNewState:=FALSE;
				_Reset();
			END_IF
			(* Check if a valid Oper_req was received *)
			IF bOperReq THEN
				bOperReq:=FALSE;
				(* Go to next ControlState *)
				_eControlState:=E_DirectControlState.PerformTest;
				bNewState:=TRUE;
			END_IF

		E_DirectControlState.PerformTest:
			(* Check if ControlState changed in the last cycle *)
			IF bNewState THEN
				bNewState:=FALSE;
				(* Set 'opRcvd' *)
				IF (_ipCtrl.ipOpRcvd <> 0) THEN
					_ipCtrl.ipOpRcvd.bValue:=TRUE;
				END_IF
			END_IF
			(* Trigger the operative test until it is finished *)
			IF _OperativeTest(bOperativeTestOk=>bTestOk, eError=>eError) THEN
				(* Reset 'opRcvd' *)
				IF (_ipCtrl.ipOpRcvd <> 0) THEN
					_ipCtrl.ipOpRcvd.bValue:=FALSE;
				END_IF
				IF bTestOk THEN
					(* Go to next ControlState *)
					_eControlState:=E_DirectControlState.WaitForExecution;
				ELSE
					fbCompletion.SetCompleted();
					fbCompletion.eServiceError:=eError;
					(* Go back to ControlState 'Ready' *)
					_eControlState:=E_DirectControlState.Ready;
				END_IF
				bNewState:=TRUE;
			END_IF

		E_DirectControlState.WaitForExecution:
			(* Check if ControlState changed in the last cycle *)
			IF bNewState THEN
				bNewState:=FALSE;
			END_IF
			(* Trigger the dynamic test until it is finished *)
			IF _DynamicTest(bDynamicTestOk=>bTestOk, eError=>eError) THEN
				fbCompletion.SetCompleted();
				IF bTestOk THEN
					(* Go to next ControlState *)
					IF (_ipBehVal <> 0) AND_THEN ((_ipBehVal.eValue = E_AcsiBeh.TestBlocked) OR_ELSE (_ipBehVal.eValue = E_AcsiBeh.OnBlocked)) THEN
						_eControlState:=E_DirectControlState.MirrorBlockedCommand;
					ELSE
						_eControlState:=E_DirectControlState.WaitForChange;
					END_IF
				ELSE
					fbCompletion.eServiceError:=eError;
					(* Go back to ControlState 'Ready' *)
					_eControlState:=E_DirectControlState.Ready;
				END_IF
				bNewState:=TRUE;
			END_IF

		E_DirectControlState.WaitForChange:
			(* Check if ControlState changed in the last cycle *)
			IF bNewState THEN
				bNewState:=FALSE;
				(* Set 'opOk' *)
				IF (_ipCtrl.ipOpOk <> 0) THEN
					_ipCtrl.ipOpOk.bValue:=TRUE;
				END_IF
				(* Set 'tOpOk' *)
				IF (_ipCtrl.ipTOpOk <> 0) AND_THEN (_ipCurrentAA <> 0) AND_THEN (_ipCurrentAA.GetSystemTime(tT=>tValue)) THEN
					_ipCtrl.ipTOpOk.tValue:=tValue;
				END_IF
			END_IF
			(* Update value *)
			_SetValue(uCtlVal:=_ipCtrl.ipOper.uCtlVal, ipCtlVal_AV:=_ipCtrl.ipOper.ipCtlVal_AnalogueValue);
			(* Update Timestamp 't' *)
			_UpdateTimestampValue(ipAA:=_ipCurrentAA);

			(* Reset 'opOk' *)
			IF (_ipCtrl.ipOpOk <> 0) THEN
				_ipCtrl.ipOpOk.bValue:=FALSE;
			END_IF
			(* Send CmdTerm_req+ *)
			_SendCommandTerminationReqPos(ipAA:=_ipCurrentAA, ipCtrlData:=_ipCtrl.ipOper);
			(* Go back to ControlState 'Ready' *)
			_eControlState:=E_DirectControlState.Ready;
			bNewState:=TRUE;

		E_DirectControlState.MirrorBlockedCommand:
			(* Check if ControlState changed in the last cycle *)
			IF bNewState THEN
				bNewState:=FALSE;
				(* Set 'opOk' *)
				IF (_ipCtrl.ipOpOk <> 0) THEN
					_ipCtrl.ipOpOk.bValue:=TRUE;
				END_IF
				(* Set 'tOpOk' *)
				IF (_ipCtrl.ipTOpOk <> 0) AND_THEN (_ipCurrentAA <> 0) AND_THEN (_ipCurrentAA.GetSystemTime(tT=>tValue)) THEN
					_ipCtrl.ipTOpOk.tValue:=tValue;
				END_IF
			END_IF
			(* Reset 'opOk' *)
			IF (_ipCtrl.ipOpOk <> 0) THEN
				_ipCtrl.ipOpOk.bValue:=FALSE;
			END_IF
			(* Send CmdTerm_req- *)
			_SendCommandTerminationReqNeg(ipAA:=_ipCurrentAA, ipCtrlData:=_ipCtrl.ipOper, eError:=E_AcsiApplError.NoError, ipOrigin:=_ipCtrl.ipOper.ipOrigin, ipCtlNum:=_ipCtrl.ipOper.ipCtlNum, eAddCause:=E_AcsiApplAddCause.BlockedByMode);
			(* Go back to ControlState 'Ready' *)
			_eControlState:=E_DirectControlState.Ready;
			bNewState:=TRUE;
	END_CASE
END_IF

(* Monitor transmission of LastApplError *)
CASE _nLastApplErrorReqState OF
	0:	;
	1:
		IF (_ipLastApplErrorReq <> 0) THEN
			Execute:=_ipLastApplErrorReq.Execute();
			IF NOT _ipLastApplErrorReq.IsBusy() THEN
				IF _ipLastApplErrorReq.IsCompleted() THEN
					SUPER^.SetCompleted();
				ELSE
					SUPER^.CopyFrom(ipSource:=_ipLastApplErrorReq);
				END_IF
				_nLastApplErrorReqState:=0;
			END_IF
		END_IF
END_CASE
(* Monitor transmission of CommandTermination *)
CASE _nCmdTermReqState OF
	0:	RETURN;
	1:
		IF (_ipCmdTermReq <> 0) THEN
			Execute:=_ipCmdTermReq.Execute();
			IF NOT _ipCmdTermReq.IsBusy() THEN
				IF _ipCmdTermReq.IsCompleted() THEN
					SUPER^.SetCompleted();
				ELSE
					SUPER^.CopyFrom(ipSource:=_ipLastApplErrorReq);
				END_IF
				_nCmdTermReqState:=0;
			END_IF
		END_IF
END_CASE
END_METHOD

END_FUNCTION_BLOCK

// ---- POUs/IEC61850Server/FB_SboControl.TcPOU
FUNCTION_BLOCK FB_SboControl EXTENDS FB_Control
VAR
	_eControlState: E_SboControlState; (*State of control state machine*)
	_fbSboTimer: TON; (*Timer to monitor 'sboTimeout'*)
END_VAR

(*This method is called when Cancel_req is received.
It shall check whether the Cancel request is valid and return FALSE as well as an error code if it is not.*)
METHOD PROTECTED _CheckCancelReq : BOOL
VAR_INPUT
	ipDai: I_AcsiDataAccessInfoClass; (*Additional data access info*)
END_VAR
VAR_OUTPUT
	eError: E_AcsiServiceError; (*Error code for negative response*)
END_VAR
VAR
	ipAA: I_ScsmAssociationClass; (*Interface pointer to application association*)
	stRemoteAddr: ST_SockAddr; (*Address of the client that sent the Cancel_req*)
END_VAR
IF (_ipCtrl <> 0) AND_THEN (_ipCtrl.ipCancel <> 0) THEN
	ScsmAssociation_From_Dai(in:=ipDai, out=>ipAA);
	(* Don't allow control if 'ctlModel' is set to 'status-only' *)
	IF (_ipCtrl.ipCtlModel <> 0) AND_THEN (_ipCtrl.ipCtlModel.eValue = E_AcsiCtlModels.StatusOnly) THEN
		_SendLastApplError(ipAA:=ipAA, ipCtrlData:=_ipCtrl.ipCancel, eError:=E_AcsiApplError.NoError, ipOrigin:=_ipCtrl.ipCancel.ipOrigin, ipCtlNum:=_ipCtrl.ipCancel.ipCtlNum, eAddCause:=E_AcsiApplAddCause.Unknown);
		RETURN;
	(* Cancel is always allowed in state 'Unselected' *)
	ELSIF (_eControlState = E_SboControlState.Unselected) THEN
		_CheckCancelReq:=TRUE;
		RETURN;
	(* Cancel is only allowed by the same client that sent the last accepted Sel_req *)
	ELSIF (RemoteAddress_From_ScsmAssociation(in:=ipAA, out=>stRemoteAddr)) AND_THEN (stRemoteAddr.sAddr <> _stCurrrentIp.sAddr) THEN
		_SendLastApplError(ipAA:=ipAA, ipCtrlData:=_ipCtrl.ipCancel, eError:=E_AcsiApplError.NoError, ipOrigin:=_ipCtrl.ipCancel.ipOrigin, ipCtlNum:=_ipCtrl.ipCancel.ipCtlNum, eAddCause:=E_AcsiApplAddCause.LockedByOtherClient);
		RETURN;
	(* Cancel is not allowed in state 'Operate' *)
	ELSIF (_eControlState = E_SboControlState.Operate) THEN
		_SendLastApplError(ipAA:=ipAA, ipCtrlData:=_ipCtrl.ipCancel, eError:=E_AcsiApplError.NoError, ipOrigin:=_ipCtrl.ipCancel.ipOrigin, ipCtlNum:=_ipCtrl.ipCancel.ipCtlNum, eAddCause:=E_AcsiApplAddCause.CommandAlreadyInExecution);
		RETURN;
	(* Cancel is valid *)
	ELSE
		_CheckCancelReq:=TRUE;
	END_IF
END_IF
END_METHOD

//Resets all local values
METHOD PROTECTED _Reset
VAR
END_VAR
SUPER^._Reset();
(* Reset timer *)
_fbSboTimer(IN:=FALSE);
END_METHOD

METHOD Execute : BOOL
VAR
	bTestOk: BOOL; (*Used to cache the return value of the last '_OperativeTest' or '_DynamicTest' method call*)
	eError: E_AcsiServiceError; (*Used to cache the returned error of the last '_OperativeTest' or '_DynamicTest' method call*)
	tValue: T_UtcTime; (*Used to cache the current system time for 'tOpOk'*)
END_VAR
IF (_ipCtrl <> 0) AND_THEN (_ipCtrl.ipOper <> 0) THEN
	(* Initialize function block in the first cycle *)
	IF NOT bInit THEN
		_Init();
		bInit:=TRUE;
	END_IF

	CASE _eControlState OF
		E_SboControlState.Unselected:
			(* Check if ControlState changed in the last cycle *)
			IF bNewState THEN
				bNewState:=FALSE;
				_Reset();
				(* Reset 'stSeld' *)
				IF (_ipCtrl.ipStSeld <> 0) THEN
					_ipCtrl.ipStSeld.bValue:=FALSE;
				END_IF
			END_IF
			(* Check if a valid Cancel_req was received *)
			IF bCancelReq THEN
				bCancelReq:=FALSE;
			END_IF
			(* Check if a valid Sel_req was received *)
			IF bSelReq THEN
				bSelReq:=FALSE;
				(* Set 'stSeld' *)
				IF (_ipCtrl.ipStSeld <> 0) THEN
					_ipCtrl.ipStSeld.bValue:=TRUE;
				END_IF
				(* Go to next ControlState *)
				_eControlState:=E_SboControlState.Ready;
				bNewState:=TRUE;
			END_IF

		E_SboControlState.Ready:
			(* Check if ControlState changed in the last cycle *)
			IF bNewState THEN
				bNewState:=FALSE;
				(* Start timer *)
				IF (_ipCtrl.ipSboTimeout <> 0) THEN
					_fbSboTimer(IN:=TRUE, PT:=DWORD_TO_TIME(_ipCtrl.ipSboTimeout.nValue));
				END_IF
			END_IF
			_fbSboTimer();
			(* Check if a valid Cancel_req was received, 'sboTimeout' was exceeded or the association was lost *)
			IF bCancelReq OR_ELSE _fbSboTimer.Q OR_ELSE ((_ipCurrentAA <> 0) AND_THEN (_ipCurrentAA.eState <> E_AsyncEnvironmentState.Established)) THEN
				bCancelReq:=FALSE;
				_fbSboTimer(IN:=FALSE);
				(* Go to next ControlState *)
				_eControlState:=E_SboControlState.EndSelection;
				bNewState:=TRUE;
			END_IF
			(* Check if a valid Oper_req was received *)
			IF bOperReq THEN
				bOperReq:=FALSE;
				(* Go to next ControlState *)
				_eControlState:=E_SboControlState.PerformTest;
				bNewState:=TRUE;
			END_IF

		E_SboControlState.PerformTest:
			(* Check if ControlState changed in the last cycle *)
			IF bNewState THEN
				bNewState:=FALSE;
				(* Set 'opRcvd' *)
				IF (_ipCtrl.ipOpRcvd <> 0) THEN
					_ipCtrl.ipOpRcvd.bValue:=TRUE;
				END_IF
			END_IF
			(* Check if a valid Cancel_req was received *)
			IF bCancelReq THEN
				bCancelReq:=FALSE;
				(* Send Oper_resp- *)
				_SendLastApplError(ipAA:=_ipCurrentAA, ipCtrlData:=_ipCtrl.ipOper, eError:=E_AcsiApplError.NoError, ipOrigin:=_ipCtrl.ipOper.ipOrigin, ipCtlNum:=_ipCtrl.ipOper.ipCtlNum, eAddCause:=E_AcsiApplAddCause.AbortionByCancel);
				fbOperCompletion.SetCompleted();
				fbOperCompletion.eServiceError:=E_AcsiServiceError.AccessViolation;
				(* Go to ControlState 'EndSelection' *)
				_eControlState:=E_SboControlState.EndSelection;
				bNewState:=TRUE;
			END_IF
			(* Trigger the operative test until it is finished *)
			IF _OperativeTest(bOperativeTestOk=>bTestOk, eError=>eError) THEN
				(* Reset 'opRcvd' *)
				IF (_ipCtrl.ipOpRcvd <> 0) THEN
					_ipCtrl.ipOpRcvd.bValue:=FALSE;
				END_IF
				IF bTestOk THEN
					(* Go to next ControlState *)
					_eControlState:=E_SboControlState.WaitForExecution;
				ELSE
					fbOperCompletion.SetCompleted();
					fbOperCompletion.eServiceError:=eError;
					(* Go to ControlState 'EndSelection' *)
					_eControlState:=E_SboControlState.EndSelection;
				END_IF
				bNewState:=TRUE;
			END_IF

		E_SboControlState.WaitForExecution:
			(* Check if ControlState changed in the last cycle *)
			IF bNewState THEN
				bNewState:=FALSE;
			END_IF
			(* Check if a Cancel_req was received *)
			IF bCancelReq THEN
				bCancelReq:=FALSE;
				(* Send Oper_resp- *)
				_SendLastApplError(ipAA:=_ipCurrentAA, ipCtrlData:=_ipCtrl.ipOper, eError:=E_AcsiApplError.NoError, ipOrigin:=_ipCtrl.ipOper.ipOrigin, ipCtlNum:=_ipCtrl.ipOper.ipCtlNum, eAddCause:=E_AcsiApplAddCause.AbortionByCancel);
				fbOperCompletion.SetCompleted();
				fbOperCompletion.eServiceError:=E_AcsiServiceError.AccessViolation;
				(* Go to ControlState 'EndSelection' *)
				_eControlState:=E_SboControlState.EndSelection;
				bNewState:=TRUE;
			END_IF
			(* Trigger the dynamic test until it is finished *)
			IF _DynamicTest(bDynamicTestOk=>bTestOk, eError=>eError) THEN
				fbOperCompletion.SetCompleted();
				IF bTestOk THEN
					(* Go to next ControlState *)
					IF (_ipBehVal <> 0) AND_THEN ((_ipBehVal.eValue = E_AcsiBeh.TestBlocked) OR_ELSE (_ipBehVal.eValue = E_AcsiBeh.OnBlocked)) THEN
						_eControlState:=E_SboControlState.MirrorBlockedCommand;
					ELSE
						_eControlState:=E_SboControlState.Operate;
					END_IF
				ELSE
					fbOperCompletion.eServiceError:=eError;
					(* Go to ControlState 'EndSelection' *)
					_eControlState:=E_SboControlState.EndSelection;
				END_IF
				bNewState:=TRUE;
			END_IF

		E_SboControlState.Operate:
			(* Check if ControlState changed in the last cycle *)
			IF bNewState THEN
				bNewState:=FALSE;
				(* Set 'opOk' *)
				IF (_ipCtrl.ipOpOk <> 0) THEN
					_ipCtrl.ipOpOk.bValue:=TRUE;
				END_IF
				(* Set 'tOpOk' *)
				IF (_ipCtrl.ipTOpOk <> 0) AND_THEN (_ipCurrentAA <> 0) AND_THEN (_ipCurrentAA.GetSystemTime(tT=>tValue)) THEN
					_ipCtrl.ipTOpOk.tValue:=tValue;
				END_IF
			END_IF
			(* Update value *)
			_SetValue(uCtlVal:=_ipCtrl.ipOper.uCtlVal, ipCtlVal_AV:=_ipCtrl.ipOper.ipCtlVal_AnalogueValue);
			(* Update Timestamp 't' *)
			_UpdateTimestampValue(ipAA:=_ipCurrentAA);

			(* Reset 'opOk' *)
			IF (_ipCtrl.ipOpOk <> 0) THEN
				_ipCtrl.ipOpOk.bValue:=FALSE;
			END_IF
			(* Go to next ControlState *)
			IF (_ipCtrl.ipSboClass <> 0) AND_THEN (_ipCtrl.ipSboClass.eValue = E_AcsiSboClasses.OperateMany) THEN
				_eControlState:=E_SboControlState.Ready;
			ELSE
				_eControlState:=E_SboControlState.EndSelection;
			END_IF
			bNewState:=TRUE;

		E_SboControlState.MirrorBlockedCommand:
			(* Check if ControlState changed in the last cycle *)
			IF bNewState THEN
				bNewState:=FALSE;
				(* Set 'opOk' *)
				IF (_ipCtrl.ipOpOk <> 0) THEN
					_ipCtrl.ipOpOk.bValue:=TRUE;
				END_IF
				(* Set 'tOpOk' *)
				IF (_ipCtrl.ipTOpOk <> 0) AND_THEN (_ipCurrentAA <> 0) AND_THEN (_ipCurrentAA.GetSystemTime(tT=>tValue)) THEN
					_ipCtrl.ipTOpOk.tValue:=tValue;
				END_IF
			END_IF
			(* Reset 'opOk' *)
			IF (_ipCtrl.ipOpOk <> 0) THEN
				_ipCtrl.ipOpOk.bValue:=FALSE;
			END_IF
			(* Go to next ControlState *)
			IF (_ipCtrl.ipSboClass <> 0) AND_THEN (_ipCtrl.ipSboClass.eValue = E_AcsiSboClasses.OperateMany) THEN
				_eControlState:=E_SboControlState.Ready;
			ELSE
				_eControlState:=E_SboControlState.EndSelection;
			END_IF
			bNewState:=TRUE;

		E_SboControlState.EndSelection:
			(* Check if ControlState changed in the last cycle *)
			IF bNewState THEN
				bNewState:=FALSE;
				(* Reset 'stSeld' *)
				IF (_ipCtrl.ipStSeld <> 0) THEN
					_ipCtrl.ipStSeld.bValue:=FALSE;
				END_IF
			END_IF
			(* Go to next ControlState *)
			_eControlState:=E_SboControlState.Unselected;
			bNewState:=TRUE;
	END_CASE
END_IF

(* Monitor transmission of LastApplError *)
CASE _nLastApplErrorReqState OF
	0:	RETURN;
	1:
		IF (_ipLastApplErrorReq <> 0) THEN
			Execute:=_ipLastApplErrorReq.Execute();
			IF NOT _ipLastApplErrorReq.IsBusy() THEN
				IF _ipLastApplErrorReq.IsCompleted() THEN
					SUPER^.SetCompleted();
				ELSE
					SUPER^.CopyFrom(ipSource:=_ipLastApplErrorReq);
				END_IF
				_nLastApplErrorReqState:=0;
			END_IF
		END_IF
END_CASE
END_METHOD

METHOD OnCompletionWaitEvent : BOOL
VAR_INPUT
	ipDai: I_AcsiDataAccessInfoClass;
	ipData: I_AcsiCommonDataClass;
	eFc: E_AcsiFc;
END_VAR
VAR_OUTPUT
	ipResult: I_AcsiServiceResultClass := fbCompletion;
END_VAR
VAR
	eServiceError: E_AcsiServiceError;
	ipAA: I_ScsmAssociationClass; (*Interface pointer to application association*)
END_VAR
fbCompletion.SetCompleted();
IF (ipDai = 0) OR_ELSE (ipData = 0) THEN
	fbCompletion.eServiceError:=E_AcsiServiceError.AccessViolation;
	RETURN;
END_IF

(* Check if an Operate request is received *)
IF (ipDai.eService = E_AcsiServiceType.SetDataValues) THEN
	IF	(ipData.sObjectName = 'Oper') THEN
		ScsmAssociation_From_Dai(in:=ipDai, out=>_ipCurrentAA);
		fbOperCompletion.SetBusy();
		ipResult:=fbOperCompletion;
		bOperReq:=TRUE;
		OnCompletionWaitEvent:=TRUE;
	ELSIF (ipData.sObjectName = 'Cancel') THEN
		fbCancelCompletion.SetCompleted();
		ipResult:=fbCancelCompletion;
		IF _CheckCancelReq(ipDai:=ipDai, eError=>eServiceError) THEN
			bCancelReq:=TRUE;
		ELSE
			fbCancelCompletion.eServiceError:=eServiceError;
		END_IF
	END_IF
END_IF
END_METHOD

(*Implementation of user application data update event method.*)
METHOD OnGetVEvent
VAR_INPUT
	ipDai: I_AcsiDataAccessInfoClass; (*Additional data access info*)
	ipData: I_AcsiCommonDataClass; (*Interface pointer to data object*)
	eFc: E_AcsiFc; (*Functional constraint*)
END_VAR
VAR
END_VAR
IF (eFc = E_AcsiFc.CO) AND_THEN (_ipCtrl <> 0) AND_THEN (ipDai <> 0) AND_THEN (ipDai.Read) AND_THEN (ipDai.ipAccessData <> 0) THEN
	IF (ipDai.ipAccessData.sObjectName = 'SBO') AND_THEN (_ipCtrl.ipSBO <> 0) THEN
		(* Reset value of 'SBO' *)
		_ipCtrl.ipSBO.sValue:='';
	END_IF
END_IF
END_METHOD

(*Implementation of user application data update event method.*)
METHOD OnGetVPreEvent : E_AcsiServiceError
VAR_INPUT
	ipDai: I_AcsiDataAccessInfoClass; (*Additional data access info*)
	ipData: I_AcsiCommonDataClass; (*Interface pointer to data object*)
	eFc: E_AcsiFc; (*Functional constraint*)
END_VAR
VAR
END_VAR
IF (eFc = E_AcsiFc.CO) AND_THEN (_ipCtrl <> 0) AND_THEN (ipDai <> 0) AND_THEN (ipDai.Read) AND_THEN (ipDai.ipAccessData <> 0) THEN
	IF (ipDai.ipAccessData.sObjectName = 'SBO') AND_THEN (_ipCtrl.ipSBO <> 0) THEN
		(* Only allow 'Select' requests in state 'Unselected' *)
		IF (_eControlState = E_SboControlState.Unselected) THEN
			_ipCtrl.ipSBO.sValue:=_ipCtrl.ipSBO.GetSboReference();
			bSelReq:=TRUE;
		ELSE
			_ipCtrl.ipSBO.sValue:='';
		END_IF
	END_IF
END_IF
END_METHOD

(*Implementation of user application data update event method.*)
METHOD OnSetVPreEvent : E_AcsiServiceError
VAR_INPUT
	ipDai: I_AcsiDataAccessInfoClass; (*Additional data access info*)
	ipMemory: I_AnyMemoryBuffer; (*Interface pointer to buffer containig new value data*)
	ipData: I_AcsiCommonDataClass; (*Interface pointer to data object*)
	eFc: E_AcsiFc; (*Functional constraint*)
END_VAR
VAR_OUTPUT
	ipLastApplError: I_AcsiDATypeLastApplError; (*IF <> 0 => send LastApplError request*)
END_VAR
VAR
	ipAA: I_ScsmAssociationClass; (*Interface pointer to application association*)
	bItself: BOOL; (*If TRUE => Checking object is sub-data object itself*)
END_VAR
IF (eFc = E_AcsiFc.CO) AND_THEN (_ipCtrl <> 0) AND_THEN (ipDai <> 0) AND_THEN (ipDai.Write) AND_THEN (ipDai.ipAccessData <> 0) AND_THEN (ipData <> 0) AND_THEN ScsmAssociation_From_Dai(in:=ipDai, out=>ipAA) THEN
	IF (_ipCtrl.ipOper <> 0) AND_THEN (_ipCtrl.ipOper.ipOrigin <> 0) AND_THEN (_ipCtrl.ipOper.ipCtlNum <> 0) THEN
		(* Check for invalid write attemps to prevent 'Oper' from being overwritten while a control request is being executed *)
		IF (ipDai.ipAccessData.sObjectName = 'Oper') THEN
			(* Only allow 'Oper' requests in state 'Ready' *)
			IF (_eControlState <> E_SboControlState.Ready) THEN
				ipLastApplError:=ipAA.SetAdditionalCauseDiag(ipCtrlData:=_ipCtrl.ipOper, eError:=E_AcsiApplError.NoError, stOrigin:=_ipCtrl.ipOper.ipOrigin.stOrigin, nCtlNum:=_ipCtrl.ipOper.ipCtlNum.nValue, eAddCause:=E_AcsiApplAddCause.CommandAlreadyInExecution);
				OnSetVPreEvent:=E_AcsiServiceError.AccessViolation;
				RETURN;
			END_IF
		ELSIF (_ipCtrl.ipOper.HasDataSubObject(ipData:=ipDai.ipAccessData, bItself=>bItself) AND_THEN (NOT bItself)) THEN
			(* Don't allow write access to subdata of 'Oper'*)
			ipLastApplError:=ipAA.SetAdditionalCauseDiag(ipCtrlData:=_ipCtrl.ipOper, eError:=E_AcsiApplError.NoError, stOrigin:=_ipCtrl.ipOper.ipOrigin.stOrigin, nCtlNum:=_ipCtrl.ipOper.ipCtlNum.nValue, eAddCause:=E_AcsiApplAddCause.NotSupported);
			OnSetVPreEvent:=E_AcsiServiceError.AccessViolation;
			RETURN;
		END_IF
	END_IF
	IF (_ipCtrl.ipCancel <> 0) AND_THEN (_ipCtrl.ipCancel.ipOrigin <> 0) AND_THEN (_ipCtrl.ipCancel.ipCtlNum <> 0) THEN
		IF (ipDai.ipAccessData.sObjectName <> 'Cancel') AND_THEN (_ipCtrl.ipCancel.HasDataSubObject(ipData:=ipDai.ipAccessData)) THEN
			(* Don't allow write access to subdata of 'Cancel'*)
			ipLastApplError:=ipAA.SetAdditionalCauseDiag(ipCtrlData:=_ipCtrl.ipCancel, eError:=E_AcsiApplError.NoError, stOrigin:=_ipCtrl.ipCancel.ipOrigin.stOrigin, nCtlNum:=_ipCtrl.ipCancel.ipCtlNum.nValue, eAddCause:=E_AcsiApplAddCause.NotSupported);
			OnSetVPreEvent:=E_AcsiServiceError.AccessViolation;
			RETURN;
		END_IF
	END_IF
	IF (ipData.sObjectName = 'SBO') THEN
		(* Don't allow write access to 'SBO'*)
		OnSetVPreEvent:=E_AcsiServiceError.AccessViolation;
		RETURN;
	END_IF
END_IF
END_METHOD

END_FUNCTION_BLOCK

// ---- POUs/IEC61850Server/FB_SboControlEnhanced.TcPOU
FUNCTION_BLOCK FB_SboControlEnhanced EXTENDS FB_SboControl
VAR
END_VAR

METHOD Execute : BOOL
VAR
	bTestOk: BOOL; (*Used to cache the return value of the last '_OperativeTest' or '_DynamicTest' method call*)
	eError: E_AcsiServiceError; (*Used to cache the returned error of the last '_OperativeTest' or '_DynamicTest' method call*)
	tValue: T_UtcTime; (*Used to cache the current system time for 'tOpOk'*)
END_VAR
IF (_ipCtrl <> 0) AND_THEN (_ipCtrl.ipOper <> 0) THEN
	(* Initialize function block in the first cycle *)
	IF NOT bInit THEN
		_Init();
		bInit:=TRUE;
	END_IF

	CASE _eControlState OF
		E_SboControlState.Unselected:
			(* Check if ControlState changed in the last cycle *)
			IF bNewState THEN
				bNewState:=FALSE;
				_Reset();
			END_IF
			(* Check if a valid Cancel_req was received *)
			IF bCancelReq THEN
				bCancelReq:=FALSE;
			END_IF
			(* Check if a valid SelVal_req was received *)
			IF bSelValReq THEN
				bSelValReq:=FALSE;
				(* Go to next ControlState *)
				_eControlState:=E_SboControlState.Select_PerformTest;
				bNewState:=TRUE;
			END_IF

		E_SboControlState.Select_PerformTest:
			(* Check if ControlState changed in the last cycle *)
			IF bNewState THEN
				bNewState:=FALSE;
			END_IF
			(* Trigger the test until it is finished *)
			IF _Test(bTestOk=>bTestOk, eError=>eError) THEN
				IF bTestOk THEN
					(* Go to next ControlState *)
					_eControlState:=E_SboControlState.WaitForSelection;
				ELSE
					fbSelValCompletion.SetCompleted();
					fbSelValCompletion.eServiceError:=eError;
					(* Go back to ControlState 'Unselected' *)
					_eControlState:=E_SboControlState.Unselected;
				END_IF
				bNewState:=TRUE;
			END_IF

		E_SboControlState.WaitForSelection:
			(* Check if ControlState changed in the last cycle *)
			IF bNewState THEN
				bNewState:=FALSE;
			END_IF
			(* Set 'stSeld' *)
			IF (_ipCtrl.ipStSeld <> 0) THEN
				_ipCtrl.ipStSeld.bValue:=TRUE;
			END_IF
			fbSelValCompletion.SetCompleted();
			(* Go to next ControlState *)
			_eControlState:=E_SboControlState.Ready;
			bNewState:=TRUE;

		E_SboControlState.Ready:
			(* Check if ControlState changed in the last cycle *)
			IF bNewState THEN
				bNewState:=FALSE;
				(* Start timer *)
				IF (_ipCtrl.ipSboTimeout <> 0) THEN
					_fbSboTimer(IN:=TRUE, PT:=DWORD_TO_TIME(_ipCtrl.ipSboTimeout.nValue));
				END_IF
			END_IF
			_fbSboTimer();
			(* Check if a valid Cancel_req was received, 'sboTimeout' was exceeded or the association was lost *)
			IF bCancelReq OR_ELSE _fbSboTimer.Q OR_ELSE ((_ipCurrentAA <> 0) AND_THEN (_ipCurrentAA.eState <> E_AsyncEnvironmentState.Established)) THEN
				bCancelReq:=FALSE;
				_fbSboTimer(IN:=FALSE);
				(* Go to next ControlState *)
				_eControlState:=E_SboControlState.EndSelection;
				bNewState:=TRUE;
			END_IF
			(* Check if a valid Oper_req was received *)
			IF bOperReq THEN
				bOperReq:=FALSE;
				(* Go to next ControlState *)
				_eControlState:=E_SboControlState.PerformTest;
				bNewState:=TRUE;
			END_IF

		E_SboControlState.PerformTest:
			(* Check if ControlState changed in the last cycle *)
			IF bNewState THEN
				bNewState:=FALSE;
				(* Set 'opRcvd' *)
				IF (_ipCtrl.ipOpRcvd <> 0) THEN
					_ipCtrl.ipOpRcvd.bValue:=TRUE;
				END_IF
			END_IF
			(* Check if a valid Cancel_req was received *)
			IF bCancelReq THEN
				bCancelReq:=FALSE;
				(* Send Oper_resp- *)
				_SendLastApplError(ipAA:=_ipCurrentAA, ipCtrlData:=_ipCtrl.ipOper, eError:=E_AcsiApplError.NoError, ipOrigin:=_ipCtrl.ipOper.ipOrigin, ipCtlNum:=_ipCtrl.ipOper.ipCtlNum, eAddCause:=E_AcsiApplAddCause.AbortionByCancel);
				fbOperCompletion.SetCompleted();
				fbOperCompletion.eServiceError:=E_AcsiServiceError.AccessViolation;
				(* Go to ControlState 'EndSelection' *)
				_eControlState:=E_SboControlState.EndSelection;
				bNewState:=TRUE;
			END_IF
			(* Trigger the operative test until it is finished *)
			IF _OperativeTest(bOperativeTestOk=>bTestOk, eError=>eError) THEN
				(* Reset 'opRcvd' *)
				IF (_ipCtrl.ipOpRcvd <> 0) THEN
					_ipCtrl.ipOpRcvd.bValue:=FALSE;
				END_IF
				IF bTestOk THEN
					(* Go to next ControlState *)
					_eControlState:=E_SboControlState.WaitForExecution;
				ELSE
					fbOperCompletion.SetCompleted();
					fbOperCompletion.eServiceError:=eError;
					(* Go to ControlState 'EndSelection' *)
					_eControlState:=E_SboControlState.EndSelection;
				END_IF
				bNewState:=TRUE;
			END_IF

		E_SboControlState.WaitForExecution:
			(* Check if ControlState changed in the last cycle *)
			IF bNewState THEN
				bNewState:=FALSE;
			END_IF
			(* Check if a Cancel_req was received *)
			IF bCancelReq THEN
				bCancelReq:=FALSE;
				(* Send Oper_resp- *)
				_SendLastApplError(ipAA:=_ipCurrentAA, ipCtrlData:=_ipCtrl.ipOper, eError:=E_AcsiApplError.NoError, ipOrigin:=_ipCtrl.ipOper.ipOrigin, ipCtlNum:=_ipCtrl.ipOper.ipCtlNum, eAddCause:=E_AcsiApplAddCause.AbortionByCancel);
				fbOperCompletion.SetCompleted();
				fbOperCompletion.eServiceError:=E_AcsiServiceError.AccessViolation;
				(* Go to ControlState 'EndSelection' *)
				_eControlState:=E_SboControlState.EndSelection;
				bNewState:=TRUE;
			END_IF
			(* Trigger the dynamic test until it is finished *)
			IF _DynamicTest(bDynamicTestOk=>bTestOk, eError=>eError) THEN
				fbOperCompletion.SetCompleted();
				IF bTestOk THEN
					(* Go to next ControlState *)
					IF (_ipBehVal <> 0) AND_THEN ((_ipBehVal.eValue = E_AcsiBeh.TestBlocked) OR_ELSE (_ipBehVal.eValue = E_AcsiBeh.OnBlocked)) THEN
						_eControlState:=E_SboControlState.MirrorBlockedCommand;
					ELSE
						_eControlState:=E_SboControlState.WaitForChange;
					END_IF
				ELSE
					fbOperCompletion.eServiceError:=eError;
					(* Go to ControlState 'EndSelection' *)
					_eControlState:=E_SboControlState.EndSelection;
				END_IF
				bNewState:=TRUE;
			END_IF

		E_SboControlState.WaitForChange:
			(* Check if ControlState changed in the last cycle *)
			IF bNewState THEN
				bNewState:=FALSE;
				(* Set 'opOk' *)
				IF (_ipCtrl.ipOpOk <> 0) THEN
					_ipCtrl.ipOpOk.bValue:=TRUE;
				END_IF
				(* Set 'tOpOk' *)
				IF (_ipCtrl.ipTOpOk <> 0) AND_THEN (_ipCurrentAA <> 0) AND_THEN (_ipCurrentAA.GetSystemTime(tT=>tValue)) THEN
					_ipCtrl.ipTOpOk.tValue:=tValue;
				END_IF
			END_IF
			(* Update value *)
			_SetValue(uCtlVal:=_ipCtrl.ipOper.uCtlVal, ipCtlVal_AV:=_ipCtrl.ipOper.ipCtlVal_AnalogueValue);
			(* Update Timestamp 't' *)
			_UpdateTimestampValue(ipAA:=_ipCurrentAA);

			(* Reset 'opOk' *)
			IF (_ipCtrl.ipOpOk <> 0) THEN
				_ipCtrl.ipOpOk.bValue:=FALSE;
			END_IF
			(* Send CmdTerm_req+ *)
			_SendCommandTerminationReqPos(ipAA:=_ipCurrentAA, ipCtrlData:=_ipCtrl.ipOper);
			(* Go to next ControlState *)
			IF (_ipCtrl.ipSboClass <> 0) AND_THEN (_ipCtrl.ipSboClass.eValue = E_AcsiSboClasses.OperateMany) THEN
				_eControlState:=E_SboControlState.Ready;
			ELSE
				_eControlState:=E_SboControlState.EndSelection;
			END_IF
			bNewState:=TRUE;

		E_SboControlState.MirrorBlockedCommand:
			(* Check if ControlState changed in the last cycle *)
			IF bNewState THEN
				bNewState:=FALSE;
				(* Set 'opOk' *)
				IF (_ipCtrl.ipOpOk <> 0) THEN
					_ipCtrl.ipOpOk.bValue:=TRUE;
				END_IF
				(* Set 'tOpOk' *)
				IF (_ipCtrl.ipTOpOk <> 0) AND_THEN (_ipCurrentAA <> 0) AND_THEN (_ipCurrentAA.GetSystemTime(tT=>tValue)) THEN
					_ipCtrl.ipTOpOk.tValue:=tValue;
				END_IF
			END_IF
			(* Reset 'opOk' *)
			IF (_ipCtrl.ipOpOk <> 0) THEN
				_ipCtrl.ipOpOk.bValue:=FALSE;
			END_IF
			(* Send CmdTerm_req- *)
			_SendCommandTerminationReqNeg(ipAA:=_ipCurrentAA, ipCtrlData:=_ipCtrl.ipOper, eError:=E_AcsiApplError.NoError, ipOrigin:=_ipCtrl.ipOper.ipOrigin, ipCtlNum:=_ipCtrl.ipOper.ipCtlNum, eAddCause:=E_AcsiApplAddCause.BlockedByMode);
			(* Go to next ControlState *)
			IF (_ipCtrl.ipSboClass <> 0) AND_THEN (_ipCtrl.ipSboClass.eValue = E_AcsiSboClasses.OperateMany) THEN
				_eControlState:=E_SboControlState.Ready;
			ELSE
				_eControlState:=E_SboControlState.EndSelection;
			END_IF
			bNewState:=TRUE;

		E_SboControlState.EndSelection:
			(* Check if ControlState changed in the last cycle *)
			IF bNewState THEN
				bNewState:=FALSE;
				(* Reset 'stSeld' *)
				IF (_ipCtrl.ipStSeld <> 0) THEN
					_ipCtrl.ipStSeld.bValue:=FALSE;
				END_IF
			END_IF
			(* Go to next ControlState *)
			_eControlState:=E_SboControlState.Unselected;
			bNewState:=TRUE;
	END_CASE
END_IF

(* Monitor transmission of LastApplError *)
CASE _nLastApplErrorReqState OF
	0:	;
	1:
		IF (_ipLastApplErrorReq <> 0) THEN
			Execute:=_ipLastApplErrorReq.Execute();
			IF NOT _ipLastApplErrorReq.IsBusy() THEN
				IF _ipLastApplErrorReq.IsCompleted() THEN
					SUPER^.SetCompleted();
				ELSE
					SUPER^.CopyFrom(ipSource:=_ipLastApplErrorReq);
				END_IF
				_nLastApplErrorReqState:=0;
			END_IF
		END_IF
END_CASE
(* Monitor transmission of CommandTermination *)
CASE _nCmdTermReqState OF
	0:	RETURN;
	1:
		IF (_ipCmdTermReq <> 0) THEN
			Execute:=_ipCmdTermReq.Execute();
			IF NOT _ipCmdTermReq.IsBusy() THEN
				IF _ipCmdTermReq.IsCompleted() THEN
					SUPER^.SetCompleted();
				ELSE
					SUPER^.CopyFrom(ipSource:=_ipLastApplErrorReq);
				END_IF
				_nCmdTermReqState:=0;
			END_IF
		END_IF
END_CASE
END_METHOD

METHOD OnCompletionWaitEvent : BOOL
VAR_INPUT
	ipDai: I_AcsiDataAccessInfoClass;
	ipData: I_AcsiCommonDataClass;
	eFc: E_AcsiFc;
END_VAR
VAR_OUTPUT
	ipResult: I_AcsiServiceResultClass := fbCompletion;
END_VAR
VAR
	eServiceError: E_AcsiServiceError;
	ipAA: I_ScsmAssociationClass; (*Interface pointer to application association*)
END_VAR
fbCompletion.SetCompleted();
IF (ipDai = 0) OR_ELSE (ipData = 0) THEN
	fbCompletion.eServiceError:=E_AcsiServiceError.AccessViolation;
	RETURN;
END_IF

(* Check if an Operate request is received *)
IF (ipDai.eService = E_AcsiServiceType.SetDataValues) THEN
	IF	(ipData.sObjectName = 'Oper') THEN
		fbOperCompletion.SetBusy();
		ipResult:=fbOperCompletion;
		bOperReq:=TRUE;
		OnCompletionWaitEvent:=TRUE;
	ELSIF (ipData.sObjectName = 'SBOw') THEN
		ScsmAssociation_From_Dai(in:=ipDai, out=>_ipCurrentAA);
		fbSelValCompletion.SetBusy();
		ipResult:=fbSelValCompletion;
		bSelValReq:=TRUE;
		OnCompletionWaitEvent:=TRUE;
	ELSIF (ipData.sObjectName = 'Cancel') THEN
		fbCancelCompletion.SetCompleted();
		ipResult:=fbCancelCompletion;
		IF _CheckCancelReq(ipDai:=ipDai, eError=>eServiceError) THEN
			bCancelReq:=TRUE;
		ELSE
			fbCancelCompletion.eServiceError:=eServiceError;
		END_IF
	END_IF
END_IF
END_METHOD

(*Implementation of user application data update event method.*)
METHOD OnGetVEvent
VAR_INPUT
	ipDai: I_AcsiDataAccessInfoClass; (*Additional data access info*)
	ipData: I_AcsiCommonDataClass; (*Interface pointer to data object*)
	eFc: E_AcsiFc; (*Functional constraint*)
END_VAR
VAR
END_VAR
END_METHOD

(*Implementation of user application data update event method.*)
METHOD OnGetVPreEvent : E_AcsiServiceError
VAR_INPUT
	ipDai: I_AcsiDataAccessInfoClass; (*Additional data access info*)
	ipData: I_AcsiCommonDataClass; (*Interface pointer to data object*)
	eFc: E_AcsiFc; (*Functional constraint*)
END_VAR
VAR
END_VAR
END_METHOD

(*Implementation of user application data update event method.*)
METHOD OnSetVPreEvent : E_AcsiServiceError
VAR_INPUT
	ipDai: I_AcsiDataAccessInfoClass; (*Additional data access info*)
	ipMemory: I_AnyMemoryBuffer; (*Interface pointer to buffer containig new value data*)
	ipData: I_AcsiCommonDataClass; (*Interface pointer to data object*)
	eFc: E_AcsiFc; (*Functional constraint*)
END_VAR
VAR_OUTPUT
	ipLastApplError: I_AcsiDATypeLastApplError; (*IF <> 0 => send LastApplError request*)
END_VAR
VAR
	ipAA: I_ScsmAssociationClass; (*Interface pointer to application association*)
	bItself: BOOL; (*If TRUE => Checking object is sub-data object itself*)
END_VAR
IF (eFc = E_AcsiFc.CO) AND_THEN (_ipCtrl <> 0) AND_THEN (ipDai <> 0) AND_THEN (ipDai.Write) AND_THEN (ipDai.ipAccessData <> 0) AND_THEN (ipData <> 0)
AND_THEN ScsmAssociation_From_Dai(in:=ipDai, out=>ipAA) THEN
	IF (_ipCtrl.ipOper <> 0) AND_THEN (_ipCtrl.ipOper.ipOrigin <> 0) AND_THEN (_ipCtrl.ipOper.ipCtlNum <> 0) THEN
		(* Check for invalid write attemps to prevent 'Oper' from being overwritten while a control request is being executed *)
		IF (ipDai.ipAccessData.sObjectName = 'Oper') THEN
			(* Only allow 'Oper' requests in state 'Ready' *)
			IF (_eControlState <> E_SboControlState.Ready) THEN
				ipLastApplError:=ipAA.SetAdditionalCauseDiag(ipCtrlData:=_ipCtrl.ipOper, eError:=E_AcsiApplError.NoError, stOrigin:=_ipCtrl.ipOper.ipOrigin.stOrigin, nCtlNum:=_ipCtrl.ipOper.ipCtlNum.nValue, eAddCause:=E_AcsiApplAddCause.CommandAlreadyInExecution);
				OnSetVPreEvent:=E_AcsiServiceError.AccessViolation;
				RETURN;
			END_IF
		ELSIF (_ipCtrl.ipOper.HasDataSubObject(ipData:=ipDai.ipAccessData, bItself=>bItself) AND_THEN (NOT bItself)) THEN
			(* Don't allow write access to subdata of 'Oper'*)
			ipLastApplError:=ipAA.SetAdditionalCauseDiag(ipCtrlData:=_ipCtrl.ipOper, eError:=E_AcsiApplError.NoError, stOrigin:=_ipCtrl.ipOper.ipOrigin.stOrigin, nCtlNum:=_ipCtrl.ipOper.ipCtlNum.nValue, eAddCause:=E_AcsiApplAddCause.NotSupported);
			OnSetVPreEvent:=E_AcsiServiceError.AccessViolation;
			RETURN;
		END_IF
	END_IF
	IF (_ipCtrl.ipSBOw <> 0) AND_THEN (_ipCtrl.ipSBOw.ipOrigin <> 0) AND_THEN (_ipCtrl.ipSBOw.ipCtlNum <> 0) THEN
		(* Check for invalid write attemps to prevent 'SBOw' from being overwritten while a control request is being executed *)
		IF (ipDai.ipAccessData.sObjectName = 'SBOw') THEN
			(* Only allow 'SelectWithValue' requests in state 'Unselected' *)
			IF (_eControlState <> E_SboControlState.Unselected) THEN
				ipLastApplError:=ipAA.SetAdditionalCauseDiag(ipCtrlData:=_ipCtrl.ipSBOw, eError:=E_AcsiApplError.NoError, stOrigin:=_ipCtrl.ipSBOw.ipOrigin.stOrigin, nCtlNum:=_ipCtrl.ipSBOw.ipCtlNum.nValue, eAddCause:=E_AcsiApplAddCause.CommandAlreadyInExecution);
				OnSetVPreEvent:=E_AcsiServiceError.AccessViolation;
				RETURN;
			ELSIF (_ipCtrl.ipSBOw.HasDataSubObject(ipData:=ipDai.ipAccessData, bItself=>bItself) AND_THEN (NOT bItself)) THEN
				(* Don't allow write access to subdata of 'SBOw'*)
				ipLastApplError:=ipAA.SetAdditionalCauseDiag(ipCtrlData:=_ipCtrl.ipSBOw, eError:=E_AcsiApplError.NoError, stOrigin:=_ipCtrl.ipSBOw.ipOrigin.stOrigin, nCtlNum:=_ipCtrl.ipSBOw.ipCtlNum.nValue, eAddCause:=E_AcsiApplAddCause.NotSupported);
				OnSetVPreEvent:=E_AcsiServiceError.AccessViolation;
				RETURN;
			END_IF
		END_IF
	END_IF
	IF (_ipCtrl.ipCancel <> 0) AND_THEN (_ipCtrl.ipCancel.ipOrigin <> 0) AND_THEN (_ipCtrl.ipCancel.ipCtlNum <> 0) THEN
		IF (ipDai.ipAccessData.sObjectName <> 'Cancel') AND_THEN (_ipCtrl.ipCancel.HasDataSubObject(ipData:=ipDai.ipAccessData)) THEN
			(* Don't allow write access to subdata of 'Cancel'*)
			ipLastApplError:=ipAA.SetAdditionalCauseDiag(ipCtrlData:=_ipCtrl.ipCancel, eError:=E_AcsiApplError.NoError, stOrigin:=_ipCtrl.ipCancel.ipOrigin.stOrigin, nCtlNum:=_ipCtrl.ipCancel.ipCtlNum.nValue, eAddCause:=E_AcsiApplAddCause.NotSupported);
			OnSetVPreEvent:=E_AcsiServiceError.AccessViolation;
			RETURN;
		END_IF
	END_IF
END_IF
END_METHOD

END_FUNCTION_BLOCK

// ---- POUs/IEC61850Server/User61850Enums/FB_ClrOp.TcPOU
{attribute 'no_explicit_call' := 'Direct call not allowed for type FB_ClrOp'}
{attribute 'call_after_init'}
FUNCTION_BLOCK FB_ClrOp EXTENDS FB_AcsiBATypeENUMERATED
VAR
	_eValue: E_ClrOp;
	_eConfig: E_ClrOp;
	{attribute 'hide'}
	ipInit: I_AcsiCommonAttributeClass := THIS^.AddDAValue(eP:=E_AcsiP.Actual, in:=_eValue).AddDAValue(eP:=E_AcsiP.Config, in:=_eConfig).AddDAType(in:=THIS^.T(in:=E_AcsiBasicType.INT8));
END_VAR

PROPERTY eConfig : E_ClrOp
GET
eConfig:= _eConfig;
END_GET
END_PROPERTY

PROPERTY eValue : E_ClrOp
GET
eValue:= _eValue;
OnGetVPropEvt();
END_GET
SET
_bChanged:= _eValue <> eValue;
_eValue:= eValue;
OnSetVPropEvt(bChanged := _bChanged);
END_SET
END_PROPERTY

END_FUNCTION_BLOCK

// ---- POUs/IEC61850Server/User61850Enums/FB_CtlMd.TcPOU
{attribute 'no_explicit_call' := 'Direct call not allowed for type FB_CtlMd'}
{attribute 'call_after_init'}
FUNCTION_BLOCK FB_CtlMd EXTENDS FB_AcsiBATypeENUMERATED
VAR
	_eValue: E_CtlMd;
	_eConfig: E_CtlMd;
	{attribute 'hide'}
	ipInit: I_AcsiCommonAttributeClass := THIS^.AddDAValue(eP:=E_AcsiP.Actual, in:=_eValue).AddDAValue(eP:=E_AcsiP.Config, in:=_eConfig).AddDAType(in:=THIS^.T(in:=E_AcsiBasicType.INT8));
END_VAR

PROPERTY eConfig : E_CtlMd
GET
eConfig:= _eConfig;
END_GET
END_PROPERTY

PROPERTY eValue : E_CtlMd
GET
eValue:= _eValue;
OnGetVPropEvt();
END_GET
SET
_bChanged:= _eValue <> eValue;
_eValue:= eValue;
OnSetVPropEvt(bChanged := _bChanged);
END_SET
END_PROPERTY

END_FUNCTION_BLOCK

// ---- POUs/IEC61850Server/User61850Enums/FB_TurCtl.TcPOU
{attribute 'no_explicit_call' := 'Direct call not allowed for type FB_TurCtl'}
{attribute 'call_after_init'}
FUNCTION_BLOCK FB_TurCtl EXTENDS FB_AcsiBATypeENUMERATED
VAR
	_eValue: E_TurCtl;
	_eConfig: E_TurCtl;
	{attribute 'hide'}
	ipInit: I_AcsiCommonAttributeClass := THIS^.AddDAValue(eP:=E_AcsiP.Actual, in:=_eValue).AddDAValue(eP:=E_AcsiP.Config, in:=_eConfig).AddDAType(in:=THIS^.T(in:=E_AcsiBasicType.INT8));
END_VAR

PROPERTY eConfig : E_TurCtl
GET
eConfig:= _eConfig;
END_GET
END_PROPERTY

PROPERTY eValue : E_TurCtl
GET
eValue:= _eValue;
OnGetVPropEvt();
END_GET
SET
_bChanged:= _eValue <> eValue;
_eValue:= eValue;
OnSetVPropEvt(bChanged := _bChanged);
END_SET
END_PROPERTY

END_FUNCTION_BLOCK
